(* IEC 61131-3 sources: daoli-st-library/DL_Process (part 68) *)

(* ---- FB_DL_MultiZoneSetpointScheduler.st ---- *)
(*==============================================================================
 * 组件名称 (Component)  : FB_DL_MultiZoneSetpointScheduler
 * 所属子库 (Sublibrary) : DL_Process ｜ 版本 (Version) : 1.0.2 ｜ 2026-11-23
 * 兼容性   (Platform)   : CODESYS 3.5+ / TwinCAT 3 / 汇川 InoProShop / 施耐德 Machine Expert
 *                         仅依赖 IEC 61131-3 标准（FOR / CASE / ABS），零厂商私有库
 * 功能描述 (Function)   : 多区设定值按时段表切换（4 区 × 每区最多 8 时段）。每区持有一张
 *                         「起始分钟 + 设定值」时段表，按当日第几分钟 nMinuteOfDay 选出生效
 *                         时段，并把「与上一生效值不同」的区以 abSpChanged 单拍沿上报。
 *                         参数非法（时段非单调 / 分钟越域 / 设定值非有限 / 时段数越界）→
 *                         整机进 eFault 并锁存首个成因码；eFault 唯一出口为 bReset（重校验通过）。
 *                         **时钟来源声明**：本件不读任何系统时钟（零全局耦合 R1），
 *                         nMinuteOfDay 由上层 PRG 从 RTC 换算后传入（0..1439）。
 *                         **bEnable = FALSE 语义（R191 二选一，本件选「冻结保持末值」）**：
 *                         各区 afActiveSp / aiActiveIdx 保持末值不动，abSpChanged 不再发沿，
 *                         bValid 落 FALSE 提示「该值已不与时钟对齐」。
 * 接口     (Interface)  : 输入 bEnable / bReset / nMinuteOfDay / aiZoneSlotCount[1..4] /
 *                         aSlots[1..4][1..8]（ST_DL_SpSlot）；输出 afActiveSp[1..4] /
 *                         aiActiveIdx[1..4] / abSpChanged[1..4]（单拍）/ eState / bError /
 *                         eCause / bValid / nFaultZone。
 * 状态迁移表 (State Transition Table)：
 *   ① eIdle → eApply：bEnable 上升（或上电首拍 bEnable 已为 TRUE）；
 *      拍 N 进入（bEnable 为 TRUE）/ 本拍行为：不做选段、不发沿、冻结保持 / 拍 N+1 转出至 eApply。
 *      拒收：bEnable 为 FALSE 时本拍不迁出，abSpChanged 保持 FALSE。
 *   ② eApply → eHold：全量参数校验通过且选段、比对、发沿完成（同一拍内完成）；
 *      拍 N 进入（校验通过）/ 本拍行为：写出 afActiveSp/aiActiveIdx 与 abSpChanged 单拍沿 /
 *      拍 N+1 转出至 eHold。
 *   ③ eApply → eFault：任一区校验失败（时段数越界 / 分钟越域 / 时段非单调 / 设定值非有限）；
 *      拍 N 进入（校验失败）/ 本拍行为：锁存首个成因码、不写 afActiveSp（保持末值）/
 *      拍 N+1 转出至 eFault（段尾迁移闸）。
 *   ④ eHold → eApply：nMinuteOfDay 落在任一时段起点（时段边界）或 bReset 为 TRUE（强制重校验）；
 *      拍 N 进入（边界命中或复位）/ 本拍行为：交出控制权、本拍不写设定值 / 拍 N+1 转出至 eApply。
 *   ⑤ eHold → eIdle：bEnable 落 FALSE（失能退出，出口冻结保持）。
 *   ⑥ eHold → eFault：段尾迁移闸（锁存位已置）——由①②③④ 任一分支置锁存后同拍迁入。
 *   ⑦ eFault → eIdle：bReset 上升且 NOT bEnable（复位沿要求先失能，避免带故障参数直接投产）；
 *      拍 N 进入（bReset 沿 + 已失能）/ 本拍行为：清锁存与成因码 / 拍 N+1 转出至 eIdle。
 *      该路径可达性自证：bReset 与 bEnable 均为外部引脚，恒可到达（R152）。
 *   ⑧ ELSE（非法枚举值）→ eFault，成因码 eIllegalState（R6 兜底）。
 * 边界     (Boundary)   : ① 首时段之前（nMinuteOfDay < 第 1 段起始）：取第 1 段值（日头承接），
 *                            该口径在段 4 注释内声明，不置码。
 *                         ② nMinuteOfDay 越域（<0 或 >1439）→ 钳位到 [0,1439] 并置信息级
 *                            eMinuteClamped（信息级永不置 bError）。
 *                         ③ 数组下标访问前先以 nCnt ∈ [1,8] 钳定（R4），越界槽不访问。
 *                         ④ 浮点同值比较用容差 DL_MZS_EPS（1E-6），禁 `=`（R4）。
 *                         ⑤ 零全局耦合（无 GVL / VAR_EXTERNAL / %I / %Q）。
 * 码表     (Codes)      : 本件不占用全局数字码位（R297 零码位范式）；出口为 BOOL + ENUM，
 *                         enum E_DL_MzsCause 归属本文件（全库唯一属主）。信息级
 *                         eMinuteClamped / eNoChange 永不置 bError；故障级成因码各占独立成员
 *                         （R190 归因唯一），锁存回放至 bReset 沿（FB33-1）。
 * 分工声明 (Scope)      : 时段选择与下发归本件；设定值斜坡 / 无扰切换归 FB_DL_RampGenerator 类；
 *                         PID 闭环归温控件。本件不下装任何硬件输出。
 * 归属     (Ownership)  : E_DL_MzsState / E_DL_MzsCause / ST_DL_SpSlot 归属本文件
 *                         （全库唯一定义，R264），引用件只引用不重声明。
 * 红线自检 (Redline)    : R1 ✓ 零 GVL ｜ R2 ✓ 零 %I/%Q ｜ R3 ✓ 纯 IEC ｜ R4 ✓ 下标钳定 +
 *                         非有限双判 + 容差比较 + 循环界固定 ｜ R5 ✓ 逐行同行双语注释
 *                         R6 ✓ 四态 ENUM + CASE + ELSE ｜ R7 N/A（本件无需定时器/边沿实例）
 *                         R14 ✓ 无 PROPERTY ｜ R8/R9 N/A（无 METHOD）
 * 修订历史 (Revision)   : 2026-11-24  v1.0.2  R79-F2/P3：bReset 电平→R_TRIG 沿 + eHold 复位沿同步清锁存（原头版本号滞留 1.0.0，已核正）
 *                         2026-11-23  v1.0.0  R78-B3 首版
 *                         2026-11-23  v1.0.1  R78 返修：E045 数组访问改嵌套索引形式（8 处）；
 *                                             eHold 相补时段数重校验闸（越界锁存 eBadCount）；
 *                                             M5：成功路径不再覆盖钳位信息级码
 * 验收向量 (Acceptance) :
 *   V1 bEnable=TRUE、nMinuteOfDay=480、区 1 时段表 {(0,20.0),(480,22.0)} → afActiveSp[1]=22.0,
 *      aiActiveIdx[1]=2, abSpChanged[1]=TRUE 单拍；次拍 abSpChanged[1]=FALSE。
 *   V2 续 V1、nMinuteOfDay 保持 481（非边界）→ eState=eHold，无沿。
 *   V3 区 2 时段表起始分钟 {0, 600, 500}（非单调）→ eState=eFault, eCause=eSlotNotMonotonic,
 *      bError=TRUE, afActiveSp[2] 保持末值；bReset 上升且 bEnable=FALSE → 回 eIdle。
 *   V4 nMinuteOfDay=2000（越域）→ 钳位到 1439，eCause=eMinuteClamped（信息级），bError=FALSE。
 *   V5 区 3 设定值为 NaN → eState=eFault, eCause=eBadSetpoint, bError=TRUE。
 *============================================================================*)

(*-----------------------------------------------------------------------------
 * 结构体: ST_DL_SpSlot（时段表行：起始分钟 + 该时段设定值），归属本文件，全库唯一属主
 *----------------------------------------------------------------------------*)
TYPE ST_DL_SpSlot :
STRUCT
    nStartMin : INT := 0;      // 时段起始时刻（当日第几分钟，0..1439）[-] / Slot start minute of the day
    fSetpoint : REAL := 0.0;   // 该时段生效设定值 [工程单位，由调用方标定] / Setpoint effective within the slot
END_STRUCT
END_TYPE

(*-----------------------------------------------------------------------------
 * 枚举: E_DL_MzsState（状态机相位；eFault 为安全相，仅 bReset 沿迁出）
 *----------------------------------------------------------------------------*)
TYPE E_DL_MzsState :
(
    eIdle  := 0,    // 空闲：未使能，设定值冻结保持末值 / Idle: disabled, setpoints frozen at last value
    eApply := 10,   // 校验与应用：全量参数校验 + 选段 + 比对 + 发沿（同拍完成）/ Validate and apply in one scan
    eHold  := 20,   // 驻留：等时段边界或复位，每拍只做边界检测 / Hold: wait for a slot boundary or reset
    eFault := 90    // 故障安全相：参数非法，锁存成因码，仅 bReset 沿迁出 / Fault latched, reset edge only
);
END_TYPE

(*-----------------------------------------------------------------------------
 * 枚举: E_DL_MzsCause（成因码；信息级 = 0..9，故障级 = 10 起，各成因独立成员 R190）
 *----------------------------------------------------------------------------*)
TYPE E_DL_MzsCause :
(
    eNone             := 0,   // 信息级：无事件 / Info: no event
    eMinuteClamped    := 1,   // 信息级：当日分钟越域已钳位 / Info: minute of day clamped into range
    eSlotNotMonotonic := 10,  // 故障级：时段起始分钟非严格递增 / Fault: slot start minutes not strictly increasing
    eBadMinute        := 11,  // 故障级：单条时段起始分钟越域 / Fault: slot start minute out of range
    eBadCount         := 12,  // 故障级：时段数越界（不在 1..8）/ Fault: slot count out of the 1..8 range
    eBadSetpoint      := 13,  // 故障级：设定值非有限 / Fault: non-finite setpoint
    eIllegalState     := 14   // 故障级：非法状态枚举值（CASE ELSE 兜底）/ Fault: illegal state enum value
);
END_TYPE

FUNCTION_BLOCK FB_DL_MultiZoneSetpointScheduler
VAR_INPUT
    bEnable        : BOOL := FALSE;                       // 使能：FALSE 冻结保持末值（本件语义声明）/ Enable, FALSE freezes the last setpoints
    bReset         : BOOL := FALSE;                       // 复位（上升沿）：清故障锁存并要求失能 / Reset rising edge clears the fault latch and requires disabled state
    nMinuteOfDay   : INT := 0;                            // 当日第几分钟，有效域 0..1439 [-] / Minute of the day, valid domain 0..1439
    aiZoneSlotCount : ARRAY[1..4] OF INT;                 // 各区时段条数，有效域 1..8 [-] / Slot count per zone, valid domain 1..8
    aSlots         : ARRAY[1..4] OF ARRAY[1..8] OF ST_DL_SpSlot;  // 四区 × 八时段时段表 / Slot tables of four zones with up to eight slots each
END_VAR
VAR_OUTPUT
    afActiveSp  : ARRAY[1..4] OF REAL;      // 各区当前生效设定值（冻结保持，见 bEnable 语义）[工程单位] / Active setpoint per zone
    aiActiveIdx : ARRAY[1..4] OF INT;       // 各区当前生效时段序号（1..8），未选定时为 0 [-] / Active slot index per zone
    abSpChanged : ARRAY[1..4] OF BOOL;      // 各区设定值变更单拍沿（统一出口预置，FB51-8）[-] / Single-scan change flag per zone
    eState      : E_DL_MzsState;            // 状态出口（段尾单点映射）[-] / State outlet, mapped at the tail
    bError      : BOOL;                     // 故障锁存标志（仅故障级成因置位）[-] / Fault latch flag
    eCause      : E_DL_MzsCause;            // 成因码出口（锁存回放）[-] / Cause code outlet, replayed from the latch
    bValid      : BOOL;                     // 设定值有效回执（eHold 且参数有效才 TRUE）[-] / Setpoint validity receipt
    nFaultZone  : INT;                      // 首个故障所在区号（0 = 无故障 / 全局性故障）[-] / Zone index of the first fault
END_VAR
VAR
    _eState      : E_DL_MzsState := E_DL_MzsState.eIdle;   // 内部相位（CASE 唯一写入目标）[-] / Internal phase
    _bFaultLatch : BOOL := FALSE;                          // 故障锁存位（仅 bReset 沿清除）[-] / Fault latch bit cleared by the reset edge only
    _eCauseLatch : E_DL_MzsCause := E_DL_MzsCause.eNone;    // 锁存成因码（锁存回放，FB33-1）[-] / Latched cause code replayed to the outlet
    _nFaultZone  : INT := 0;                               // 首个故障区号 [1..4]，0 表示无 / Zone index of the first fault
    _bParamOk    : BOOL := TRUE;                           // 本拍参数校验通过标志 [-] / Parameter validation flag of this scan
    _eCauseTmp   : E_DL_MzsCause := E_DL_MzsCause.eNone;    // 本拍首个成因（未锁存）[-] / First cause of this scan before latching
    _nFaultZtmp  : INT := 0;                               // 本拍首个故障区号（未锁存）[-] / First fault zone of this scan before latching
    _nMinute     : INT := 0;                               // 钳位后的当日分钟 [0..1439] / Clamped minute of the day
    _nCnt        : INT := 0;                               // 当前区时段条数（校验后使用）[-] / Slot count of the current zone
    _nIdx        : INT := 0;                               // 选段中间结果（时段序号）[-] / Intermediate slot index
    _nNewIdx     : INT := 0;                               // 本区本拍应生效时段序号 [-] / Slot index that should be active this scan
    _fNewSp      : REAL := 0.0;                            // 本区本拍应生效设定值 [工程单位] / Setpoint that should be active this scan
    _bBoundary   : BOOL := FALSE;                          // 时段边界命中标志（eHold 用）[-] / Slot boundary hit flag used in eHold
    _nZ          : INT := 0;                               // 外层循环索引：区号 [1..4] / Outer loop index, zone number
    _nK          : INT := 0;                               // 内层循环索引：时段序号 [1..8] / Inner loop index, slot number
    _rtReset     : R_TRIG;                                 // 复位沿检测实例（v1.0.1 补：声明沿即实现沿，段 1 无条件刷新）/ Reset edge detector, refreshed unconditionally in segment 1
END_VAR
VAR CONSTANT
    DL_MZS_ZONES    : INT := 4;             // 固定区数（数组第一维上界）[-] / Fixed zone count, upper bound of dimension one
    DL_MZS_SLOTS    : INT := 8;             // 每区最大时段数（数组第二维上界）[-] / Max slots per zone, upper bound of dimension two
    DL_MZS_MIN_DAY  : INT := 1439;          // 当日最大分钟数（23:59）[-] / Last minute of the day
    DL_MZS_MIN_ONE  : INT := 1;             // 时段数下界 [-] / Lower bound of the slot count
    DL_MZS_ZERO     : INT := 0;             // 整数零基准 [-] / Integer zero base
    DL_MZS_FZERO    : REAL := 0.0;          // 实数零基准 [-] / Real zero base
    DL_MZS_EPS      : REAL := 1.0E-6;       // 设定值同值判定容差 [-] / Setpoint equality tolerance
    DL_MZS_FIN      : LREAL := 1.0E308;     // 有限性判据上界（R477：ABS(x)>FIN 判 Inf）[工程单位] / finiteness ceiling flags Inf
END_VAR

(* —— 段 1：单拍位与当拍工作量预置（只清单拍标志，不清锁存/保持量，FB32-1） —— *)
_rtReset(CLK := bReset);                                // 复位沿刷新必须无条件周期调用（R7；v1.0.1 修复 J1 电平判据缺陷）/ The reset edge must be refreshed unconditionally every scan
FOR _nZ := 1 TO DL_MZS_ZONES DO
    abSpChanged[_nZ] := FALSE;                          // 变更沿每拍先预清 / Change edge preset FALSE every scan
END_FOR
_bParamOk   := TRUE;                                    // 校验标志复位 / Validation flag reset
_eCauseTmp  := E_DL_MzsCause.eNone;                      // 当拍成因复位 / Scan cause reset
_nFaultZtmp := DL_MZS_ZERO;                             // 当拍故障区复位 / Scan fault zone reset
_bBoundary  := FALSE;                                   // 边界标志复位 / Boundary flag reset
eCause      := E_DL_MzsCause.eNone;                      // 成因出口每拍预置信息级零码（段 2/段 3 内改写）/ Cause outlet preset to the info zero code every scan

(* —— 段 2：入参钳位与域闸（分钟越域钳位并置信息级，R4 下标与域安全） —— *)
_nMinute := nMinuteOfDay;                               // 取入参 / Take the input pin
IF _nMinute < DL_MZS_ZERO THEN
    _nMinute  := DL_MZS_ZERO;                           // 下越界钳到 0 / Clamp low
    eCause    := E_DL_MzsCause.eMinuteClamped;          // 信息级：已钳位 / Info: clamped
ELSIF _nMinute > DL_MZS_MIN_DAY THEN
    _nMinute  := DL_MZS_MIN_DAY;                        // 上越界钳到 1439 / Clamp high
    eCause    := E_DL_MzsCause.eMinuteClamped;          // 信息级：已钳位 / Info: clamped
END_IF

(* —— 段 3：状态机主体（唯一相位写入点，每分支迁移条件自足） —— *)
CASE _eState OF
    E_DL_MzsState.eIdle :
        (* 迁移①：使能上升进入统一校验相；未使能则保持冻结语义 *)
        IF bEnable THEN
            _eState := E_DL_MzsState.eApply;            // 迁入校验与应用相 / Move to validate-and-apply
        END_IF

    E_DL_MzsState.eApply :
        IF NOT bEnable THEN
            _eState := E_DL_MzsState.eIdle;             // 使能消失：退回冻结 / Enable gone: back to idle
        ELSE
            (* 段 4 前置：逐区全量校验（时段数 → 单条分钟 → 单调性 → 设定值有限性） *)
            FOR _nZ := 1 TO DL_MZS_ZONES DO
                _nCnt := aiZoneSlotCount[_nZ];          // 取本区时段条数 / Slot count of this zone
                IF (_nCnt < DL_MZS_MIN_ONE) OR (_nCnt > DL_MZS_SLOTS) THEN
                    _bParamOk := FALSE;                 // 时段数越界 / Count out of range
                    IF _eCauseTmp = E_DL_MzsCause.eNone THEN
                        _eCauseTmp  := E_DL_MzsCause.eBadCount;    // 首因锁存用 / First cause kept
                        _nFaultZtmp := _nZ;                        // 记录故障区号 / Record the fault zone
                    END_IF
                ELSE
                    FOR _nK := 1 TO _nCnt DO
                        (* 单条起始分钟域闸：0..1439 *)
                        IF (aSlots[_nZ][_nK].nStartMin < DL_MZS_ZERO)
                            OR (aSlots[_nZ][_nK].nStartMin > DL_MZS_MIN_DAY) THEN
                            _bParamOk := FALSE;
                            IF _eCauseTmp = E_DL_MzsCause.eNone THEN
                                _eCauseTmp  := E_DL_MzsCause.eBadMinute;   // 故障级：分钟越域
                                _nFaultZtmp := _nZ;
                            END_IF
                        END_IF
                        (* 单调性闸：自第 2 条起必须严格大于前一条 *)
                        IF _nK > 1 THEN
                            IF aSlots[_nZ][_nK].nStartMin <= aSlots[_nZ][_nK - 1].nStartMin THEN
                                _bParamOk := FALSE;
                                IF _eCauseTmp = E_DL_MzsCause.eNone THEN
                                    _eCauseTmp  := E_DL_MzsCause.eSlotNotMonotonic;   // 故障级：非单调
                                    _nFaultZtmp := _nZ;
                                END_IF
                            END_IF
                        END_IF
                        (* 设定值有限性闸（R79 双判） *)
                        (* v1.0.2 补（闸 Q2）：Inf 判据改 R477 范式 ABS(x) > DL_MZS_FIN，
                           x−x 差判在部分编译器会常量折叠成 0，Inf 设定值可穿透写入 afActiveSp *)
                        IF (aSlots[_nZ][_nK].fSetpoint <> aSlots[_nZ][_nK].fSetpoint)
                            OR (ABS(aSlots[_nZ][_nK].fSetpoint) > DL_MZS_FIN) THEN
                            _bParamOk := FALSE;
                            IF _eCauseTmp = E_DL_MzsCause.eNone THEN
                                _eCauseTmp  := E_DL_MzsCause.eBadSetpoint;   // 故障级：设定值非有限
                                _nFaultZtmp := _nZ;
                            END_IF
                        END_IF
                    END_FOR
                END_IF
            END_FOR

            IF NOT _bParamOk THEN
                (* 迁移③：校验失败 → 锁存首因（不改写 afActiveSp，保持末值） *)
                _eCauseLatch := _eCauseTmp;                 // 锁存成因码 / Latch the cause code
                _nFaultZone  := _nFaultZtmp;                // 锁存故障区号 / Latch the fault zone
                _bFaultLatch := TRUE;                       // 置故障锁存（段尾迁移闸迁相）/ Latch the fault
            ELSE
                (* 段 4：选段 + 比对 + 发沿（每区独立裁决，日头承接口径见分支注释） *)
                FOR _nZ := 1 TO DL_MZS_ZONES DO
                    _nCnt   := aiZoneSlotCount[_nZ];        // 时段条数 / Slot count
                    _nNewIdx := DL_MZS_MIN_ONE;             // 缺省取第 1 段（日头承接：首段之前沿用首段值）/ Default first slot
                    FOR _nK := 1 TO _nCnt DO
                        IF aSlots[_nZ][_nK].nStartMin <= _nMinute THEN
                            _nNewIdx := _nK;                // 最后一条不晚于当前分钟的时段生效 / Last slot not later than now wins
                        END_IF
                    END_FOR
                    _fNewSp := aSlots[_nZ][_nNewIdx].fSetpoint;    // 取该时段设定值 / Setpoint of the winning slot
                    IF (ABS(afActiveSp[_nZ] - _fNewSp) >= DL_MZS_EPS) OR (aiActiveIdx[_nZ] <> _nNewIdx) THEN
                        afActiveSp[_nZ]  := _fNewSp;            // 写入生效设定值 / Write the active setpoint
                        aiActiveIdx[_nZ] := _nNewIdx;           // 写入生效时段序号 / Write the active slot index
                        abSpChanged[_nZ] := TRUE;               // 单拍变更沿（本拍置位，次拍段 1 预清）/ Single-scan change edge
                    END_IF
                END_FOR
                IF eCause <> E_DL_MzsCause.eMinuteClamped THEN
                    eCause := E_DL_MzsCause.eNone;          // 信息级：无事件（M5：不覆盖段 2 已置的钳位信息码）/ Info: no event, keep the pre-set clamp code
                END_IF
                _bFaultLatch := FALSE;                      // 校验通过：清故障锁存（正常路径唯一清点）/ Clear the latch on the valid path
                _eState := E_DL_MzsState.eHold;             // 迁移②：进入驻留相 / Move to hold
            END_IF
        END_IF

    E_DL_MzsState.eHold :
        IF NOT bEnable THEN
            _eState := E_DL_MzsState.eIdle;                 // 迁移⑤：失能退出（冻结保持）/ Disable exit, frozen
        ELSE
            (* 边界检测：任一时段起点等于当前分钟（或日切 0 点）→ 回校验相重算 *)
            IF _nMinute = DL_MZS_ZERO THEN
                _bBoundary := TRUE;                         // 日切 0 点视为边界 / Day roll-over counts as a boundary
            END_IF
            FOR _nZ := 1 TO DL_MZS_ZONES DO
                _nCnt := aiZoneSlotCount[_nZ];              // 取本区时段条数（引脚每拍可被外部改写，不信任 eApply 旧校验）/ Slot count, pin may change every scan
                IF (_nCnt < DL_MZS_MIN_ONE) OR (_nCnt > DL_MZS_SLOTS) THEN
                    (* L1 加固：eHold 相重校验失败 → 故障锁存（复用参数校验闸同款 eBadCount），跳出该区处理 *)
                    IF _eCauseLatch = E_DL_MzsCause.eNone THEN   // 首因保留（不覆盖既有锁存码）/ Keep the first cause
                        _eCauseLatch := E_DL_MzsCause.eBadCount; // 故障级：时段数越界（既有成因成员，R190）/ Fault: count out of range
                        _nFaultZone  := _nZ;                     // 锁存故障区号 / Latch the fault zone
                    END_IF
                    _bFaultLatch := TRUE;                        // 置故障锁存（段 5 迁移闸同拍迁入 eFault）/ Latch the fault
                ELSE
                    FOR _nK := 1 TO _nCnt DO
                        IF aSlots[_nZ][_nK].nStartMin = _nMinute THEN
                            _bBoundary := TRUE;                 // 时段边界命中 / Slot boundary hit
                        END_IF
                    END_FOR
                END_IF
            END_FOR
            IF _rtReset.Q THEN
                (* v1.0.2 补（闸 P3）：eHold 内复位沿属"强制重校验"语义，必须同时清故障锁存，
                   否则 eApply 重校验通过后 bError 仍为 TRUE（声明"复位即清锁存"未兑现） *)
                _bFaultLatch := FALSE;                      // 复位沿清故障锁存 / Reset edge clears the fault latch
                _eCauseLatch := E_DL_MzsCause.eNone;        // 复位沿清锁存成因 / Reset edge clears the latched cause
                eCause       := E_DL_MzsCause.eNone;        // 出口同步归零 / Outlet follows
                nFaultZone   := DL_MZS_ZERO;                // 故障区号归零 / Fault zone index cleared
            END_IF
            IF (NOT _bFaultLatch) AND (_bBoundary OR _rtReset.Q) THEN
                _eState := E_DL_MzsState.eApply;            // 迁移④：边界命中或强制重校验（R274：锁存期禁迁入执行相）/ Boundary or forced revalidation
            END_IF
        END_IF

    E_DL_MzsState.eFault :
        (* 迁移⑦：唯一出口 —— bReset 沿 + 已失能（避免带故障参数直接投产） *)
        IF _rtReset.Q AND (NOT bEnable) THEN
            _bFaultLatch := FALSE;                          // 清故障锁存 / Clear the fault latch
            _eCauseLatch := E_DL_MzsCause.eNone;            // 清锁存成因 / Clear the latched cause
            _nFaultZone  := DL_MZS_ZERO;                    // 清故障区号 / Clear the fault zone
            _eState      := E_DL_MzsState.eIdle;            // 回空闲相 / Back to idle
        END_IF

ELSE
    (* 迁移⑧：非法枚举值兜底（R6） *)
    _eCauseLatch := E_DL_MzsCause.eIllegalState;            // 故障级：非法状态 / Fault: illegal state value
    _bFaultLatch := TRUE;                                   // 置锁存 / Latch
    _eState      := E_DL_MzsState.eFault;                   // 迁入安全相 / Move to the safe state
END_CASE

(* —— 段 5：段尾故障迁移闸（FB50-1④：锁存与迁相分离，置于解除段之后） —— *)
IF _bFaultLatch AND (_eState <> E_DL_MzsState.eFault) THEN
    _eState := E_DL_MzsState.eFault;                        // 锁存即迁相 / Latch forces the fault phase
END_IF

(* —— 段 6：统一出口（状态映射 + 锁存回放 + 单拍位已由段 1 预置） —— *)
eState := _eState;                                          // 相位映射 / Phase mapping
bError := _bFaultLatch;                                     // 故障标志取锁存位（派生式）/ Fault flag derived from the latch
IF _bFaultLatch THEN
    eCause := _eCauseLatch;                                 // 故障期回放锁存码（FB33-1）/ Replay the latched code
    nFaultZone := _nFaultZone;                              // 回放故障区号 / Replay the fault zone
ELSE
    nFaultZone := DL_MZS_ZERO;                              // 无故障：区号归零 / No fault: zone index zero
END_IF
bValid := (_eState = E_DL_MzsState.eHold) AND (NOT _bFaultLatch);   // 仅驻留相且无锁存时值可信 / Valid only in hold without a latch
END_FUNCTION_BLOCK

(* ---- FB_DL_OccScheduleWindow.st ---- *)
(*==============================================================================
 * 组件名称 (Component)  : FB_DL_OccScheduleWindow
 * 所属子库 (Sublibrary) : DL_Process
 * 当前版本 (Version)    : 1.0.0
 * 组件分类 (Category)   : 功能块（FUNCTION_BLOCK）· 多窗作息排程 ·
 *                         Level 2 行业池 9.5 节 P0 链路闭环示范
 * 兼容性   (Platform)   : CODESYS 3.5 / TwinCAT 3 / 汇川 InoProShop / Schneider
 *                         Machine Expert；仅依赖 Standard.library（R_TRIG /
 *                         MIN）与本库 DL_Base 已入库组件，零厂商方言
 * 功能描述 (Function)   : 多窗作息排程块（最多 4 窗并行）。日期/时刻全部引脚
 *                         注入（零全局耦合红线：禁读 CPU 本地钟）→ 调用
 *                         FC_DL_DayOfWeekCalc 换算当日星期（ISO-8601 序）
 *                         → 内部 4 实例复用 FB_DL_TimeWindowCheck 逐窗判定
 *                         （每日窗矩阵 + 节假日覆盖位）→ 输出占用合成、
 *                         占用开始沿单发、活动窗号（多窗同开取最小号）与
 *                         预启动占位（提前启机预热/预冷用）。
 * 设计要点 (Key notes)  : ① 每窗占用 = 窗实例 bInWindow（内部已合成 总使能
 *                           AND 星期位 AND 时刻窗），总使能引脚折入
 *                           bEnableDay := aWinEnable[i] AND NOT aHoliday-
 *                           Override[i]（节假日强制当日该窗关闭）；窗实例的
 *                           aWeekdayEnable 由本块按 aWeekdayWin[i, 当日星期]
 *                           单日位展开为 7 日表填充；
 *                         ② 预启动占位：折算「占用开始时刻 − tPreLeadTime」
 *                           分钟域判定。推导：窗开始分钟 uStartMin（UINT 域，
 *                           0..1439，与 FB_DL_TimeWindowCheck 折算口径一致）；
 *                           当 提前量 ≤ 开始时刻 时预启带 = [开始−提前, 开始)
 *                           （左闭右开）；当 提前量 > 开始时刻（跨零点回绕）
 *                           时预启带 = [开始+24h−提前, 开始)∪[0, 开始)，即
 *                           [开始+1440−lead, 1440) 与 [0, 开始) 的并——本块
 *                           统一用 TIME 域表达（T#24H 回绕式），时刻折算先
 *                           USINT→DINT 扩宽再乘 60 防溢出（复用窗实例口径，
 *                           声明一致）；预启带归属注入日期当日窗（跨零点前段
 *                           归属前一日期的同一窗组态，调用方按日切换注入即可）；
 *                         ③ 窗实例与沿检测实例在主体无条件周期刷新（R7，
 *                           严禁置于 IF/CASE 分支）；
 *                         ④ 【事件型+日切换沿，免首扫（R23）】输入输出均为
 *                           电平/日历注入，无连续量同步语义，窗判定为组合
 *                           逻辑逐拍重算，故不设 bInit 首扫判据；
 *                         ⑤ 日期越界（FC 返回 eInvalid）→ 全窗按不在窗处理
 *                           + 信息级 0005_0210；各窗实例信息级码 0001_0202
 *                           不透传，本块归并为自身码 0005_0211（头注释声明）；
 *                         ⑥ bReset 上升沿清除当拍信息级码（日切换后防陈旧码
 *                           残留），不影响窗判定结果（沿用窗实例 D2 语义）；
 *                         ⑦ 本块无浮点量，非有限值防御不适用（公约 0.8 N/A）。
 * 枚举归属 (Enum note)  : 复用 E_DL_Weekday（DL_Base，随 FC_DL_DayOfWeekCalc
 *                         同文件发布的既有公开契约，直接引用，禁止重定义）；
 *                         本块不新增任何 DUT。
 * 依赖     (Depends)    : FB_DL_TimeWindowCheck（DL_Base，4 实例复用）；
 *                         FC_DL_DayOfWeekCalc + E_DL_Weekday（DL_Base）；
 *                         Standard.library：R_TRIG / MIN。
 * 开源溯源 (Origin)     : 原创实现（参考 OSCAT Building 时钟排程族与
 *                         Siemens LGF 定时开关族的公开行为定义，clean-room）。
 *                         仅借鉴「多窗排程 + 星期使能矩阵 + 节假日覆盖」的
 *                         公开行为语义；多实例单一语义组合架构、预启动占位、
 *                         时间引脚注入均为本库独立设计，未复制任何源码行。
 * 故障码表 (Error codes):
 *   16#0005_0210【信息级】日期参数越界（年/月/日，FC 返回 eInvalid），全窗
 *                 按不在窗处理
 *   16#0005_0211【信息级】窗时刻参数越界（各窗实例 0001_0202 码不透传，本块
 *                 归并为自身码；实例侧越界已钳位照常计算，本块预启动判定对
 *                 参数越界窗按跳过处理）
 *   【02xx 段信息级占位声明（规格 §7 有意裁定，R11 留档）】0210/0211 占用
 *   02xx 段：日历排程块全部事件均为信息级（无安全联锁、无锁存故障位），
 *   故障级段整体保留给后续工艺联锁件，沿用 FB_DL_TimeWindowCheck 先例，
 *   避免读者误判为故障级。
 * 红线自检 (Redline)    : R1 ✓ 零全局变量表与外部变量引用 ｜ R2 ✓ 零物理 IO 地址直写
 *                         R3 ✓ 纯 IEC 61131-3 ｜ R4 ✓ 数组索引域校验+USINT→DINT
 *                             扩宽防溢出+TIME 回绕防御（提前量钳位）；无浮点量，
 *                             非有限值防御不适用（R23 事件型）
 *                         R5 ✓ 全变量中英双语同行注释
 *                         R6 不适用（组合逻辑+沿检测，无状态机；星期换算
 *                           CASE 含 ELSE 兜底）
 *                         R7 ✓ 4 个窗实例 + 2 个 R_TRIG 实例主体无条件周期刷新
 * 修订历史 (Revision)   :
 *   2026-11-15  v1.0.0  首版入库 · Round 06 · 泳道 C · 契约出处 ROUND_PLAN_R6 §3.15
 * 验收向量 (Acceptance) :
 *   V1 单窗占用链：窗 1 On=08:00/Off=18:00 使能，Now=07:59 → bOccupied=
 *      FALSE；08:00 当拍 bPulseOnOccupy=TRUE 单发且 bOccupied=TRUE；
 *      18:00 当拍 bOccupied=FALSE（左闭右开与窗实例一致）
 *   V2 四窗并行：窗 2 与窗 4 同时在窗 → uActiveWin=2（多窗同开取最小号）
 *   V3 节假日覆盖：aHolidayOverride[1]=TRUE → 当日窗 1 强制不在窗，其余窗
 *      不受影响
 *   V4 预启动提前量（含跨零点回绕）：tPreLeadTime=T#30M，窗 On=06:00 →
 *      Now=05:35 bPreStart=TRUE 且 bOccupied=FALSE，06:00 当拍 bPreStart
 *      随占用置位而清零；跨零点窗 On=00:10、提前量 30 分 → Now=23:50 时
 *      bPreStart=TRUE（预启带 [23:40, 00:10)，回绕式 开始+24h−提前=23:40）
 *   V5 日期越界降级：uMonth=13 → FC 返回 eInvalid → 全窗不在窗 +
 *      0005_0210；bReset 沿当拍清码
 *   V6 星期矩阵按日生效：aWeekdayWin[1,6]=FALSE（周六位）→ 周六窗 1 不在窗，
 *      周一~周五正常
 *============================================================================*)

(*-----------------------------------------------------------------------------
 * 调用示例 (Instance guide)：
 *   fbOcc.uYear := 2026; fbOcc.uMonth := 11; fbOcc.uDay := 15;   // 日历注入
 *   fbOcc.uHourNow := stClock.hour; fbOcc.uMinNow := stClock.min;
 *   fbOcc.aWinEnable[1] := TRUE; fbOcc.aHourOn[1] := 8;         // 窗 1 组态，其余 3 窗同构
 *   fbOcc(tPreLeadTime := T#30M, bReset := bDaySwReset);         // 周期调用
 *   预热/预冷联动：bPreStart → AHU 通风预启（非占用占位）；bPulseOnOccupy
 *   → 占用开始沿一次性事件（照明/门禁联动）。uActiveWin 供 HMI 显示当前窗。
 *----------------------------------------------------------------------------*)

FUNCTION_BLOCK FB_DL_OccScheduleWindow
VAR_INPUT
    uYear              : UINT;             // 日期注入-年（Injected date year）[年] 有效域 1980..2099，越界返回 eInvalid（透传 FC_DL_DayOfWeekCalc）
    uMonth             : USINT;            // 日期注入-月（Injected month）[月] 有效域 1..12，越界按日期非法处理
    uDay               : USINT;            // 日期注入-日（Injected day）[日] 有效域 1..当月天数（含闰年），越界按日期非法处理
    uHourNow           : USINT;            // 当前时刻注入-时（Injected time hour）[h] 0..23，越界按不在窗处理（禁读 CPU 钟，公约 0.9）
    uMinNow            : USINT;            // 当前时刻注入-分（Injected time minute）[min] 0..59
    aWinEnable         : ARRAY[1..4] OF BOOL;          // 各窗使能（Window enables）[1] 窗 1..4，FALSE 时该窗恒不在窗
    aHourOn            : ARRAY[1..4] OF USINT;         // 各窗开启时刻-时（Window on hours）[h] 0..23，越界该窗预启动跳过（实例侧钳位照算）
    aMinOn             : ARRAY[1..4] OF USINT;         // 各窗开启时刻-分（Window on minutes）[min] 0..59
    aHourOff           : ARRAY[1..4] OF USINT;         // 各窗关闭时刻-时（Window off hours）[h] 0..23，支持跨零点窗
    aMinOff            : ARRAY[1..4] OF USINT;         // 各窗关闭时刻-分（Window off minutes）[min] 0..59
    aWeekdayWin        : ARRAY[1..4, 1..7] OF BOOL;    // 各窗星期使能矩阵（Per-window weekday matrix）[1] 第二维 1=周一..7=周日（ISO 序）
    aHolidayOverride   : ARRAY[1..4] OF BOOL;          // 节假日覆盖位（Holiday overrides）[1] TRUE=当日该窗强制关闭
    tPreLeadTime       : TIME := T#30M;    // 预启动提前量（Pre-start lead time）默认 T#30M，防御钳位 ≤ T#12H，占用开始前输出预启动占位
    bReset             : BOOL := FALSE;    // 复位（Reset）[1] 上升沿：清除当拍信息级码（不影响窗判定）
END_VAR
VAR_OUTPUT
    bOccupied          : BOOL;             // 占用中（Occupied）[1] 任一有效窗在窗内
    bPreStart          : BOOL;             // 预启动占位（Pre-start placeholder）[1] 未占用且距某有效窗开始 ≤ 提前量
    bPulseOnOccupy     : BOOL;             // 占用开始沿单发（Occupancy start edge）[1] TRUE 持续一拍
    uActiveWin         : USINT;            // 当前活动窗号（Active window index）1..4，0=无，多窗同开取最小号
    uErrorId           : UDINT;            // 信息级码（Info code）16#0005_0210 日期非法 / 16#0005_0211 窗参数越界；0 = 无
END_VAR
VAR
    _fbWin1            : FB_DL_TimeWindowCheck;  // 窗 1 判定实例（Window 1 checker instance）
    _fbWin2            : FB_DL_TimeWindowCheck;  // 窗 2 判定实例（Window 2 checker instance）
    _fbWin3            : FB_DL_TimeWindowCheck;  // 窗 3 判定实例（Window 3 checker instance）
    _fbWin4            : FB_DL_TimeWindowCheck;  // 窗 4 判定实例（Window 4 checker instance）
    fbTrigReset        : R_TRIG;                 // 复位信号上升沿检测实例（Reset edge detector）
    fbTrigOccupy       : R_TRIG;                 // 占用开始沿检测实例（Occupancy edge detector），CLK = bOccupied
    _eWd               : E_DL_Weekday := E_DL_Weekday.eInvalid;  // 星期换算返回值（Weekday calc result，复用 DL_Base 既有枚举）
    _uErrDow           : UDINT;                  // 星期换算返回码（Weekday calc code）16#0001_0201 = 日期越界
    _bDateOk           : BOOL;                   // 日期有效性（Date valid）
    _uWd               : USINT;                  // 当日星期 USINT 域（Current weekday）1..7，0=非法
    _bWdOk             : BOOL;                   // 星期索引有效性（Weekday index valid）
    _bTimeOk           : BOOL;                   // 当前时刻有效性（Time-of-day valid）
    _abWdSel           : ARRAY[1..7] OF BOOL;    // 单日位展开表（Expanded single-day table），喂窗实例 aWeekdayEnable
    abEnDay            : ARRAY[1..4] OF BOOL;    // 各窗日总使能（Per-window day enable）= 窗使能 AND NOT 节假日覆盖
    abWdBit            : ARRAY[1..4] OF BOOL;    // 各窗当日星期位（Per-window weekday bit）
    abWinValid         : ARRAY[1..4] OF BOOL;    // 各窗今日有效（Per-window valid today）= 日使能 AND 星期位 AND 开启参数合法
    abOccWin           : ARRAY[1..4] OF BOOL;    // 各窗占用结果（Per-window occupancy）
    abPreBand          : ARRAY[1..4] OF BOOL;    // 各窗预启带命中（Per-window pre-start band hit）
    _nNowMin           : DINT;                   // 当前时刻折算分钟（Now in minutes）0..1439，USINT→DINT 扩宽防溢出
    _nStartMin         : DINT;                   // 窗开始折算分钟（Start in minutes）0..1439，扩宽防溢出
    _atStartT          : ARRAY[1..4] OF TIME;    // 各窗开始时刻 TIME 域（Per-window start time），分钟折算防溢出后换域
    _tNowT             : TIME;                   // 当前时刻 TIME 域（Now in TIME domain），预启带比较用
    _tLeadT            : TIME;                   // 生效提前量（Effective lead time）防御钳位 ≤ T#12H
    _i                 : USINT;                  // 循环索引（Loop index）1..4，固定界防死循环
    _j                 : USINT;                  // 循环索引（Loop index）1..7，固定界防死循环
END_VAR

// -----------------------------------------------------------------------------
// 段 1｜复位沿实例无条件周期刷新（R7 红线：严禁移入 IF/CASE 分支）
// -----------------------------------------------------------------------------
fbTrigReset(CLK := bReset);                 // 复位沿检测

// -----------------------------------------------------------------------------
// 段 2｜出口默认值与时刻有效性（事件型逐拍重算，无状态驻留）
// -----------------------------------------------------------------------------
uErrorId := 16#0000_0000;                   // 信息级码每拍重算
bOccupied := FALSE;                         // 占用合成默认 FALSE
bPreStart := FALSE;                         // 预启动默认 FALSE
bPulseOnOccupy := FALSE;                    // 沿单发默认 FALSE（段 10 覆盖）
uActiveWin := 0;                            // 活动窗号默认无
_bTimeOk := (uHourNow <= 23) AND (uMinNow <= 59);   // 时刻域检查（越界预启动跳过）

// -----------------------------------------------------------------------------
// 段 3｜星期换算：FC_DL_DayOfWeekCalc 公开接口直接调用（不内联重实现）
// -----------------------------------------------------------------------------
_eWd := FC_DL_DayOfWeekCalc(uYear := uYear, uMonth := uMonth, uDay := uDay,
                            uErrorId => _uErrDow);              // 日期 → 星期（ISO 序）
_bDateOk := (_uErrDow = 16#0000_0000);                          // 返回码 0 = 日期合法
IF NOT _bDateOk THEN
    uErrorId := 16#0005_0210;               // 日期非法【信息级】：全窗按不在窗处理
END_IF

// 星期枚举 → USINT 索引显式映射（strict 枚举不整型直赋；CASE+ELSE 兜底）
CASE _eWd OF
    E_DL_Weekday.eMonday:    _uWd := 1;     // 周一（ISO 1）
    E_DL_Weekday.eTuesday:   _uWd := 2;     // 周二（ISO 2）
    E_DL_Weekday.eWednesday: _uWd := 3;     // 周三（ISO 3）
    E_DL_Weekday.eThursday:  _uWd := 4;     // 周四（ISO 4）
    E_DL_Weekday.eFriday:    _uWd := 5;     // 周五（ISO 5）
    E_DL_Weekday.eSaturday:  _uWd := 6;     // 周六（ISO 6）
    E_DL_Weekday.eSunday:    _uWd := 7;     // 周日（ISO 7）
    ELSE
        _uWd := 0;                          // eInvalid / 未预期：当日全窗不使能
END_CASE
_bWdOk := (_uWd >= 1) AND (_uWd <= 7);      // 索引域校验（防矩阵越界，R4）

// -----------------------------------------------------------------------------
// 段 4｜公共量预计算：日使能 / 星期位 / 窗有效性 / 开始时刻折算（分钟域扩宽）
// -----------------------------------------------------------------------------
FOR _i := 1 TO 4 DO
    abEnDay[_i] := aWinEnable[_i] AND (NOT aHolidayOverride[_i]);   // 日总使能 = 窗使能 AND NOT 节假日
    abWdBit[_i] := FALSE;                   // 星期位默认 FALSE（索引非法时全窗不使能）
    IF _bWdOk THEN
        abWdBit[_i] := aWeekdayWin[_i, _uWd];   // 当日星期位（索引 1..7 已校验）
    END_IF
    abWinValid[_i] := abEnDay[_i] AND abWdBit[_i]
                   AND (aHourOn[_i] <= 23) AND (aMinOn[_i] <= 59);
                                            // 今日有效 = 日使能 AND 星期位 AND 开启参数合法
    _nStartMin := aHourOn[_i];              // USINT → DINT 扩宽（先赋值再乘防溢出）
    _nStartMin := (_nStartMin * 60) + aMinOn[_i];   // 开窗分钟 0..1439
    _atStartT[_i] := T#1M * _nStartMin;     // 分钟域 → TIME 域（MUL(TIME, 整数) 标准序）
END_FOR

_nNowMin := uHourNow;                       // USINT → DINT 扩宽
_nNowMin := (_nNowMin * 60) + uMinNow;      // 当前分钟 0..1439（越界值仅预启带门控弃用）
_tNowT := T#1M * _nNowMin;                  // 当前时刻 → TIME 域
_tLeadT := tPreLeadTime;                    // 提前量原值生效
IF _tLeadT > T#12H THEN
    _tLeadT := T#12H;                       // 防御钳位：提前量组态域建议 ≤ 半日，回绕式防负时长
END_IF

// -----------------------------------------------------------------------------
// 段 5~8｜窗 1~4 实例逐拍无条件刷新（R7：调用与输入准备均不入 IF/CASE 分支）
//        每窗：单日位展开 → 实例调用 → 占用收集 → 实例码归并 → 预启带判定
// -----------------------------------------------------------------------------

// ---- 窗 1（Window 1）----
FOR _j := 1 TO 7 DO
    _abWdSel[_j] := abWdBit[1];             // aWeekdayWin[1, 当日] 单日位展开为 7 日表
END_FOR
_fbWin1(uHourNow := uHourNow, uMinNow := uMinNow,
        bEnableDay := abEnDay[1], aWeekdayEnable := _abWdSel, uWeekdayNow := _uWd,
        uHourOn := aHourOn[1], uMinOn := aMinOn[1],
        uHourOff := aHourOff[1], uMinOff := aMinOff[1], bReset := FALSE);
                                            // 窗 1 实例刷新（bReset 恒 FALSE：实例码仅当拍归并）
abOccWin[1] := _fbWin1.bInWindow;           // 窗 1 占用结果
IF _bDateOk AND (_fbWin1.uErrorId <> 16#0000_0000) THEN
    uErrorId := 16#0005_0211;               // 实例码不透传，归并为本块 0211【信息级】
END_IF
abPreBand[1] := FALSE;                      // 预启带默认未命中
IF abWinValid[1] AND _bTimeOk THEN
    IF _tLeadT <= _atStartT[1] THEN
        abPreBand[1] := (_tNowT >= (_atStartT[1] - _tLeadT)) AND (_tNowT < _atStartT[1]);
                                            // 同日内预启带 [开始−提前, 开始) 左闭右开
    ELSE
        abPreBand[1] := (_tNowT >= ((_atStartT[1] + T#24H) - _tLeadT))
                    OR (_tNowT < _atStartT[1]);
                                            // 跨零点回绕：预启带 [开始+24h−提前, 24h)∪[0, 开始)
    END_IF
END_IF

// ---- 窗 2（Window 2）----
FOR _j := 1 TO 7 DO
    _abWdSel[_j] := abWdBit[2];             // aWeekdayWin[2, 当日] 单日位展开
END_FOR
_fbWin2(uHourNow := uHourNow, uMinNow := uMinNow,
        bEnableDay := abEnDay[2], aWeekdayEnable := _abWdSel, uWeekdayNow := _uWd,
        uHourOn := aHourOn[2], uMinOn := aMinOn[2],
        uHourOff := aHourOff[2], uMinOff := aMinOff[2], bReset := FALSE);
                                            // 窗 2 实例刷新
abOccWin[2] := _fbWin2.bInWindow;           // 窗 2 占用结果
IF _bDateOk AND (_fbWin2.uErrorId <> 16#0000_0000) THEN
    uErrorId := 16#0005_0211;               // 实例码归并【信息级】
END_IF
abPreBand[2] := FALSE;                      // 预启带默认未命中
IF abWinValid[2] AND _bTimeOk THEN
    IF _tLeadT <= _atStartT[2] THEN
        abPreBand[2] := (_tNowT >= (_atStartT[2] - _tLeadT)) AND (_tNowT < _atStartT[2]);
                                            // 同日内预启带
    ELSE
        abPreBand[2] := (_tNowT >= ((_atStartT[2] + T#24H) - _tLeadT))
                    OR (_tNowT < _atStartT[2]);
                                            // 跨零点回绕预启带
    END_IF
END_IF

// ---- 窗 3（Window 3）----
FOR _j := 1 TO 7 DO
    _abWdSel[_j] := abWdBit[3];             // aWeekdayWin[3, 当日] 单日位展开
END_FOR
_fbWin3(uHourNow := uHourNow, uMinNow := uMinNow,
        bEnableDay := abEnDay[3], aWeekdayEnable := _abWdSel, uWeekdayNow := _uWd,
        uHourOn := aHourOn[3], uMinOn := aMinOn[3],
        uHourOff := aHourOff[3], uMinOff := aMinOff[3], bReset := FALSE);
                                            // 窗 3 实例刷新
abOccWin[3] := _fbWin3.bInWindow;           // 窗 3 占用结果
IF _bDateOk AND (_fbWin3.uErrorId <> 16#0000_0000) THEN
    uErrorId := 16#0005_0211;               // 实例码归并【信息级】
END_IF
abPreBand[3] := FALSE;                      // 预启带默认未命中
IF abWinValid[3] AND _bTimeOk THEN
    IF _tLeadT <= _atStartT[3] THEN
        abPreBand[3] := (_tNowT >= (_atStartT[3] - _tLeadT)) AND (_tNowT < _atStartT[3]);
                                            // 同日内预启带
    ELSE
        abPreBand[3] := (_tNowT >= ((_atStartT[3] + T#24H) - _tLeadT))
                    OR (_tNowT < _atStartT[3]);
                                            // 跨零点回绕预启带
    END_IF
END_IF

// ---- 窗 4（Window 4）----
FOR _j := 1 TO 7 DO
    _abWdSel[_j] := abWdBit[4];             // aWeekdayWin[4, 当日] 单日位展开
END_FOR
_fbWin4(uHourNow := uHourNow, uMinNow := uMinNow,
        bEnableDay := abEnDay[4], aWeekdayEnable := _abWdSel, uWeekdayNow := _uWd,
        uHourOn := aHourOn[4], uMinOn := aMinOn[4],
        uHourOff := aHourOff[4], uMinOff := aMinOff[4], bReset := FALSE);
                                            // 窗 4 实例刷新
abOccWin[4] := _fbWin4.bInWindow;           // 窗 4 占用结果
IF _bDateOk AND (_fbWin4.uErrorId <> 16#0000_0000) THEN
    uErrorId := 16#0005_0211;               // 实例码归并【信息级】
END_IF
abPreBand[4] := FALSE;                      // 预启带默认未命中
IF abWinValid[4] AND _bTimeOk THEN
    IF _tLeadT <= _atStartT[4] THEN
        abPreBand[4] := (_tNowT >= (_atStartT[4] - _tLeadT)) AND (_tNowT < _atStartT[4]);
                                            // 同日内预启带
    ELSE
        abPreBand[4] := (_tNowT >= ((_atStartT[4] + T#24H) - _tLeadT))
                    OR (_tNowT < _atStartT[4]);
                                            // 跨零点回绕预启带
    END_IF
END_IF

// -----------------------------------------------------------------------------
// 段 9｜占用合成与活动窗号（多窗同开取最小号；日期非法时全窗自然为 FALSE）
// -----------------------------------------------------------------------------
bOccupied := abOccWin[1] OR abOccWin[2] OR abOccWin[3] OR abOccWin[4];
                                            // 任一有效窗在窗内即占用
FOR _i := 1 TO 4 DO
    IF abOccWin[_i] AND (uActiveWin = 0) THEN
        uActiveWin := _i;                   // 取最小活动窗号（升序首中）
    END_IF
END_FOR

bPreStart := (NOT bOccupied) AND _bTimeOk
         AND (abPreBand[1] OR abPreBand[2] OR abPreBand[3] OR abPreBand[4]);
                                            // 预启动：未占用 AND 时刻合法 AND 任一有效窗预启带命中

// -----------------------------------------------------------------------------
// 段 10｜占用开始沿单发（实例无条件周期刷新，沿输出持续一拍）
// -----------------------------------------------------------------------------
fbTrigOccupy(CLK := bOccupied);             // 占用上升沿检测（主体无条件调用）
bPulseOnOccupy := fbTrigOccupy.Q;           // 占用开始沿单发输出

// -----------------------------------------------------------------------------
// 段 11｜复位沿消费：清除当拍信息级码（触发实例已在段 1 无条件刷新）
// -----------------------------------------------------------------------------
IF fbTrigReset.Q THEN
    uErrorId := 16#0000_0000;               // 复位沿当拍清信息级码（下一拍重新评估）
END_IF

END_FUNCTION_BLOCK

(* ---- FB_DL_PalletizerLayerBuildSeq.st ---- *)
(*==============================================================================
 * 组件名称 (Component)  : FB_DL_PalletizerLayerBuildSeq
 * 所属子库 (Sublibrary) : DL_Process ｜ 版本 (Version) : 1.0.2 ｜ 2026-11-23
 * 兼容性   (Platform)   : CODESYS 3.5+ / TwinCAT 3 / 汇川 InoProShop / 施耐德 Machine Expert
 *                         仅依赖 IEC 61131-3 标准库（TON 属 Standard.library），零厂商私有库
 * 功能描述 (Function)   : 码垛层构建时序：eIdle →（bStart）→ ePick（发取料指令，等
 *                         bPickDone 到位）→ ePlace（发放料指令，等 bPlaceDone 到位并计数）
 *                         → 满层判（nPlacedInLayer ≥ nBoxPerLayer）→ eLayerDone（发单拍层完成沿）
 *                         → 换层（nLayerNo + 1，层内计数清零）回 ePick；层数达 nLayersPerPallet
 *                         → eFull（整垛完成，等 bStart 跌落或复位）。取 / 放每相均带
 *                         tPhaseTimeout 超时兜底 → eFault。
 *                         **输出语义**：bPickCmd / bPlaceCmd 为电平台（相驻留期间为 TRUE），
 *                         bLayerDone 为**单拍脉冲**（内部 _bLayerDoneInt 置位 → 统一出口映射，
 *                         两段式，FB33-1），每拍由段 1 预置 FALSE，故脉冲宽度恰一扫描。
 *                         **bStart = FALSE 语义（R191 二选一，本件选「降级为安全值 + 置标志」）**：
 *                         全部动作输出落 FALSE 并回 eIdle（码垛动作不得冻结保持，冻结即撞机）。
 * 接口     (Interface)  : 输入 bStart / bReset / bPickDone / bPlaceDone / nBoxPerLayer /
 *                         nLayersPerPallet / tPhaseTimeout；输出 bPickCmd / bPlaceCmd /
 *                         nPlacedInLayer / nLayerNo / bLayerDone / bPalletFull / eState /
 *                         bError / eCause / bValid。
 * 状态迁移表 (State Transition Table)：
 *   ① eIdle → ePick：bStart 为 TRUE 且组态校验通过（nBoxPerLayer / nLayersPerPallet 均在域内）；
 *      拍 N 进入（启动）/ 本拍行为：层内计数与层号初始化（nPlacedInLayer := 0、nLayerNo := 1）、
 *      不发指令 / 拍 N+1 转出至 ePick。
 *   ② ePick → ePlace：bPickDone 上升沿（本拍事件优先于超时，FB51-5）；拍 N 进入（取料到位）/
 *      本拍行为：撤 bPickCmd、发 bPlaceCmd / 拍 N+1 转出至 ePlace。
 *   ③ ePick → eFault：tonPhase.Q（超时）；拍 N 进入（超时）/ 本拍行为：锁存 ePickTimeout、
 *      撤全部动作 / 拍 N+1 转出至 eFault（段尾迁移闸）。
 *   ④ ePlace → ePick：bPlaceDone 上升沿且层未满（nPlacedInLayer + 1 < nBoxPerLayer）；
 *      拍 N 进入（放料到位）/ 本拍行为：层内计数 +1、撤 bPlaceCmd / 拍 N+1 转出至 ePick。
 *   ⑤ ePlace → eLayerDone：bPlaceDone 上升沿且本次计数后层已满；拍 N 进入 /
 *      本拍行为：层内计数 +1、_bLayerDoneInt := TRUE / 拍 N+1 转出至 eLayerDone。
 *   ⑥ ePlace → eFault：tonPhase.Q（超时），锁存 ePlaceTimeout。
 *   ⑦ eLayerDone → eFull：nLayerNo ≥ nLayersPerPallet；拍 N 进入 / 本拍行为：bPalletFull := TRUE /
 *      拍 N+1 转出至 eFull。
 *   ⑧ eLayerDone → ePick：层未满垛；拍 N 进入 / 本拍行为：nLayerNo + 1、nPlacedInLayer := 0 /
 *      拍 N+1 转出至 ePick。
 *   ⑨ eFull → eIdle：bStart 落 FALSE（前置条件消失）或 bReset 为 TRUE（两条出口，R98）；
 *      拍 N 进入 / 本拍行为：层号与层内计数清零、bPalletFull 落 FALSE / 拍 N+1 转出至 eIdle。
 *   ⑩ eFault → eIdle：bReset 上升且 bStart 为 FALSE（可达性自证 R152：两引脚外部恒可达）；
 *      拍 N 进入 / 本拍行为：清锁存与成因 / 拍 N+1 转出至 eIdle。
 *   ⑪ ELSE（非法枚举值）→ eFault，成因 eIllegalState（R6 兜底）。
 * 边界     (Boundary)   : ① 相超时 TON 在 CASE 外无条件调用（R7 / FB50-1①），IN 表达式为
 *                            「处于取/放相 AND 相已稳定一拍（nPhase = nPhasePrev）AND
 *                            非故障相 AND 非故障锁存」——相切换那一拍 IN 为 FALSE 使 ET 自清，
 *                            结构性无需外部沿清零（R188）。
 *                         ② 组态域闸：nBoxPerLayer ∈ [1,60]、nLayersPerPallet ∈ [1,40]，
 *                            越域置故障级 eBadConfig（R4，兼作数组/计数安全）。
 *                         ③ ePick / ePlace 退出条件均为「事件沿 + 超时」两条（R98）。
 *                         ④ 无数组、无除法，故无下标与除零风险。
 *                         ⑤ 零全局耦合（无 GVL / VAR_EXTERNAL / %I / %Q）。
 * 码表     (Codes)      : 本件不占用全局数字码位（R297 零码位范式）；出口为 BOOL + ENUM，
 *                         enum E_DL_PlbCause 归属本文件（全库唯一属主）。信息级
 *                         eLayerDoneCode 永不置 bError；超时 / 组态 / 非法状态各占独立成员
 *                         （R190 归因唯一），锁存回放至 bReset 沿（FB33-1）。
 * 分工声明 (Scope)      : 层内路径规划 / 码型排布归 FB_DL_PalletizerStation 与
 *                         FB_DL_PalletizerLayerSeq（区段时序）；夹爪安全归 FB_DL_PalletGripperSafe。
 *                         本件只做「取—放—满层—换层—满垛」的计数与时序，不做轴运动与轨迹。
 * 归属     (Ownership)  : E_DL_PlbState / E_DL_PlbCause 归属本文件（全库唯一定义，R264）。
 * 红线自检 (Redline)    : R1 ✓ 零 GVL ｜ R2 ✓ 零 %I/%Q ｜ R3 ✓ 纯 IEC ｜ R4 ✓ 组态域闸 +
 *                         无除法无下标 + 计数单调 ｜ R5 ✓ 逐行同行双语注释 ｜ R6 ✓ 六态 ENUM +
 *                         CASE + ELSE ｜ R7 ✓ tonPhase 在 CASE 外无条件调用 ｜ R14 ✓ 无 PROPERTY
 *                         R8/R9 N/A（无 METHOD）｜ FB32-6 ✓ 单拍脉冲置位与撤销分属两拍
 * 修订历史 (Revision)   : 2026-11-23  v1.0.0  R78-B3 首版
 * 验收向量 (Acceptance) :
 *   V1 nBoxPerLayer=2、nLayersPerPallet=2：bStart 上升 → ePick；bPickDone 脉冲 → ePlace；
 *      bPlaceDone 脉冲 → nPlacedInLayer=1 且回 ePick；再一轮 → nPlacedInLayer=2、eLayerDone、
 *      bLayerDone 单拍为 TRUE（次拍 FALSE）；随后 nLayerNo=2、nPlacedInLayer=0、ePick。
 *   V2 续 V1 完成第 2 层 → eFull、bPalletFull=TRUE；bStart 落 FALSE → 回 eIdle，计数全清。
 *   V3 tPhaseTimeout=5s、bPickDone 始终不来 → 5s 后 eState=eFault、eCause=ePickTimeout、
 *      bError=TRUE、bPickCmd=FALSE；bReset 上升且 bStart=FALSE → 回 eIdle。
 *   V4 nBoxPerLayer=0 → eState=eFault、eCause=eBadConfig、bError=TRUE。
 *   V5 eFull 内 bReset=TRUE（bStart 仍 TRUE）→ 回 eIdle 并清计数（第二条出口）。
 *============================================================================*)

(*-----------------------------------------------------------------------------
 * 枚举: E_DL_PlbState（码垛层构建相位；eFault 为安全相，仅 bReset 沿迁出）
 *----------------------------------------------------------------------------*)
TYPE E_DL_PlbState :
(
    eIdle      := 0,    // 空闲：无动作输出，等 bStart / Idle: no motion command, waiting for bStart
    ePick      := 10,   // 取料相：bPickCmd 电平为 TRUE，等 bPickDone / Pick phase: bPickCmd high until bPickDone
    ePlace     := 20,   // 放料相：bPlaceCmd 电平为 TRUE，等 bPlaceDone / Place phase: bPlaceCmd high until bPlaceDone
    eLayerDone := 30,   // 层完成相：发 bLayerDone 单拍沿并判定换层 / Layer done: emit the single-scan edge and decide
    eFull      := 40,   // 整垛完成相：bPalletFull 电平为 TRUE / Pallet full: bPalletFull high
    eFault     := 90    // 故障安全相：超时 / 组态非法，动作全撤 / Fault safe phase: timeout or bad configuration
);
END_TYPE

(*-----------------------------------------------------------------------------
 * 枚举: E_DL_PlbCause（成因码；信息级 = 0..9，故障级 = 10 起）
 *----------------------------------------------------------------------------*)
TYPE E_DL_PlbCause :
(
    eNone          := 0,   // 信息级：无事件 / Info: no event
    eLayerDoneCode := 1,   // 信息级：一层已构建完成 / Info: one layer completed
    ePalletDone    := 2,   // 信息级：整垛完成 / Info: pallet completed
    ePickTimeout   := 10,  // 故障级：取料相超时 / Fault: pick phase timeout
    ePlaceTimeout  := 11,  // 故障级：放料相超时 / Fault: place phase timeout
    eBadConfig     := 12,  // 故障级：每层箱数 / 每垛层数越域 / Fault: box-per-layer or layer count out of domain
    eIllegalState  := 13   // 故障级：非法状态枚举值 / Fault: illegal state enum value
);
END_TYPE

FUNCTION_BLOCK FB_DL_PalletizerLayerBuildSeq
VAR_INPUT
    bStart          : BOOL := FALSE;          // 启动（电平）：FALSE 时动作全撤并回 eIdle / Start level, FALSE withdraws all commands
    bReset          : BOOL := FALSE;          // 复位（上升沿，需同时 bStart=FALSE）/ Reset rising edge, requires bStart FALSE
    bPickDone       : BOOL := FALSE;         // 取料到位反馈（上升沿表示本相完成，初值 FALSE 防首拍假沿）/ Pick completion feedback, rising edge ends the phase, FALSE default avoids a first-scan ghost edge
    bPlaceDone      : BOOL := FALSE;         // 放料到位反馈（上升沿表示本相完成，初值 FALSE 防首拍假沿）/ Place completion feedback, rising edge ends the phase, FALSE default avoids a first-scan ghost edge
    nBoxPerLayer    : INT := 5;               // 每层箱数，有效域 1..60 [-] / Boxes per layer, valid domain 1..60
    nLayersPerPallet : INT := 6;              // 每垛层数，有效域 1..40 [-] / Layers per pallet, valid domain 1..40
    tPhaseTimeout   : TIME := T#10S;          // 单相超时（取/放共用），域 > 0 [s] / Phase timeout shared by pick and place
END_VAR
VAR_OUTPUT
    bPickCmd        : BOOL;                   // 取料指令（电平）/ Pick command, level signal
    bPlaceCmd       : BOOL;                   // 放料指令（电平）/ Place command, level signal
    nPlacedInLayer  : INT := 0;               // 本层已放箱数 [个] / Boxes placed in the current layer
    nLayerNo        : INT := 0;               // 当前层号（1 起）[层] / Current layer number starting at one
    bLayerDone      : BOOL;                   // 层完成单拍脉冲（段 1 预置，统一出口映射）[-] / Single-scan layer-done pulse
    bPalletFull     : BOOL;                   // 整垛完成（电平，保持至 bStart 跌落或复位）[-] / Pallet full, level held until bStart falls or reset
    eState          : E_DL_PlbState;           // 状态出口（段尾单点映射）[-] / State outlet mapped at the tail
    bError          : BOOL;                   // 故障锁存标志 [-] / Fault latch flag
    eCause          : E_DL_PlbCause;          // 成因码出口（故障期锁存回放）[-] / Cause code outlet
    bValid          : BOOL;                   // 时序有效回执（取/放相才 TRUE）[-] / Sequence validity receipt
END_VAR
VAR
    _eState        : E_DL_PlbState := E_DL_PlbState.eIdle;    // 内部相位（CASE 唯一写入目标）[-] / Internal phase
    _eStatePrev    : E_DL_PlbState := E_DL_PlbState.eIdle;    // 上一拍相位快照（相稳定判据用，段末唯一更新）[-] / Phase snapshot of the last scan
    _bFaultLatch   : BOOL := FALSE;                           // 故障锁存位（仅 bReset 沿清除）[-] / Fault latch bit
    _eCauseLatch   : E_DL_PlbCause := E_DL_PlbCause.eNone;     // 锁存成因码（FB33-1 锁存回放）[-] / Latched cause code
    _bCfgOk        : BOOL := TRUE;                            // 组态域闸通过标志 [-] / Configuration gate flag
    _bLayerDoneInt : BOOL := FALSE;                           // 层完成内部单拍位（统一出口映射，FB33-1）[-] / Internal single-scan layer-done bit
    _bPhaseActive  : BOOL := FALSE;                           // 取/放相驻留标志（超时使能域）[-] / Phase-resident flag driving the timeout
    _bPickRise     : BOOL := FALSE;                           // 取料到位上升沿（本拍）/ Pick completion rising edge of this scan
    _bPlaceRise    : BOOL := FALSE;                           // 放料到位上升沿（本拍）/ Place completion rising edge of this scan
    rtPickDone     : R_TRIG;                                  // 取料到位边沿实例（段 3 无条件调用）/ Pick edge instance called unconditionally
    rtPlaceDone    : R_TRIG;                                  // 放料到位边沿实例（段 3 无条件调用）/ Place edge instance called unconditionally
    tonPhase       : TON;                                     // 相超时定时器（段 3 无条件调用）/ Phase timeout timer called unconditionally
    _rtReset     : R_TRIG;                                 // 复位沿检测实例（v1.0.2 补：声明沿即实现沿，CASE 外无条件刷新）/ Reset edge detector refreshed outside the CASE
END_VAR
VAR CONSTANT
    DL_PLB_ZERO      : INT := 0;      // 计数零基准 [-] / Count zero base
    DL_PLB_ONE       : INT := 1;      // 计数起始值（层号与每层首箱）[-] / Count start value
    DL_PLB_BOX_MAX   : INT := 60;     // 每层箱数上限（域闸用）[-] / Upper bound of boxes per layer
    DL_PLB_LAYER_MAX : INT := 40;     // 每垛层数上限（域闸用）[-] / Upper bound of layers per pallet
END_VAR

(* —— 段 1：单拍位与动作出口预置（纸清单拍标志与电平出口，不清锁存/计数，FB32-1） —— *)
bLayerDone     := FALSE;                                // 单拍层完成沿每拍预清 / Single-scan edge preset FALSE every scan
bPickCmd       := FALSE;                                // 取料指令预置（安全侧：默认不动作）/ Pick command preset, safe side
bPlaceCmd      := FALSE;                                // 放料指令预置（安全侧：默认不动作）/ Place command preset, safe side
_bLayerDoneInt := FALSE;                                // 内部单拍位预清 / Internal single-scan bit preset
_bCfgOk        := TRUE;                                 // 组态闸标志复位 / Configuration flag reset

(* —— 段 2：组态域闸（每层箱数 / 每垛层数，R4） —— *)
IF (nBoxPerLayer < DL_PLB_ONE) OR (nBoxPerLayer > DL_PLB_BOX_MAX)
    OR (nLayersPerPallet < DL_PLB_ONE) OR (nLayersPerPallet > DL_PLB_LAYER_MAX) THEN
    _bCfgOk := FALSE;                                   // 组态越域 / Configuration out of domain
    IF NOT _bFaultLatch THEN
        _eCauseLatch := E_DL_PlbCause.eBadConfig;       // 故障级：组态非法（首因锁存）/ Fault: bad configuration
        _bFaultLatch := TRUE;                           // 置故障锁存 / Latch the fault
    END_IF
END_IF

(* —— 段 3：边沿与超时实例（CASE 外无条件调用，R7 / FB50-1①） —— *)
rtPickDone(CLK := bPickDone);                           // 取料到位沿（无条件刷新：非取料相期间的沿被吞，属 R7 固有口径）/ Pick completion edge, refreshed unconditionally, edges outside the phase are consumed
rtPlaceDone(CLK := bPlaceDone);                         // 放料到位沿（无条件刷新，沿吞噬口径与取料沿一致）/ Place completion edge, refreshed unconditionally with the same edge-consumption rule
_bPickRise  := rtPickDone.Q;                            // 取料沿快照 / Pick edge snapshot
_bPlaceRise := rtPlaceDone.Q;                           // 放料沿快照 / Place edge snapshot
_bPhaseActive := (_eState = E_DL_PlbState.ePick) OR (_eState = E_DL_PlbState.ePlace);   // 取/放相驻留 / Phase residency
tonPhase(IN := _bPhaseActive AND (_eState = _eStatePrev) AND (_eState <> E_DL_PlbState.eFault) AND (NOT _bFaultLatch),
         PT := tPhaseTimeout);                          // 相稳定一拍后才计时，相切换拍 ET 自清（R188）/ Timer armed only after a stable phase scan

(* —— 段 4：状态机主体（唯一相位写入点，事件沿优先于超时，FB51-5） —— *)
_rtReset(CLK := bReset);                                // 复位沿刷新无条件周期调用（R7；v1.0.2 修复 J1 电平判据缺陷 / R18）/ Refresh the reset edge unconditionally every scan
CASE _eState OF
    E_DL_PlbState.eIdle :
        IF bStart AND (NOT _bFaultLatch) THEN
            nPlacedInLayer := DL_PLB_ZERO;              // 层内计数清零 / Clear the in-layer count
            nLayerNo       := DL_PLB_ONE;               // 层号置 1 / Start at layer one
            bPalletFull    := FALSE;                    // 整垛标志复位 / Clear the pallet-full flag
            eCause         := E_DL_PlbCause.eNone;      // 信息级：无事件 / Info: no event
            _eState        := E_DL_PlbState.ePick;      // 迁移①：进入取料相 / Move to pick
        ELSE
            bPalletFull := FALSE;                       // 未启动：整垛标志保持 FALSE / Not started: pallet flag FALSE
        END_IF

    E_DL_PlbState.ePick :
        bPickCmd := TRUE;                               // 取料指令电平为 TRUE / Pick command high
        IF _bPickRise THEN
            (* 迁移②：本拍事件优先，先消化到位沿再消化超时（FB51-5） *)
            bPickCmd := FALSE;                          // 撤取料指令 / Withdraw the pick command
            eCause   := E_DL_PlbCause.eNone;            // 信息级：无事件 / Info: no event
            _eState  := E_DL_PlbState.ePlace;           // 迁入放料相 / Move to place
        ELSIF tonPhase.Q THEN
            (* 迁移③：超时兜底 *)
            _eCauseLatch := E_DL_PlbCause.ePickTimeout; // 故障级：取料超时 / Fault: pick timeout
            _bFaultLatch := TRUE;                       // 置故障锁存 / Latch the fault
            bPickCmd     := FALSE;                      // 撤动作 / Withdraw the command
            _eState      := E_DL_PlbState.eFault;       // 迁入故障相 / Move to fault
        END_IF

    E_DL_PlbState.ePlace :
        bPlaceCmd := TRUE;                              // 放料指令电平为 TRUE / Place command high
        IF _bPlaceRise THEN
            (* 迁移④ / ⑤：放料到位 → 计数 + 满层判（两出口分列） *)
            bPlaceCmd      := FALSE;                    // 撤放料指令 / Withdraw the place command
            nPlacedInLayer := nPlacedInLayer + DL_PLB_ONE;   // 层内计数 +1 / Increment the in-layer count
            IF nPlacedInLayer >= nBoxPerLayer THEN
                _bLayerDoneInt := TRUE;                 // 层已满：内部单拍位置位（统一出口映射）/ Layer full: internal edge bit
                eCause         := E_DL_PlbCause.eLayerDoneCode;   // 信息级：一层完成 / Info: one layer done
                _eState        := E_DL_PlbState.eLayerDone;       // 迁入层完成相 / Move to layer done
            ELSE
                eCause := E_DL_PlbCause.eNone;          // 信息级：无事件 / Info: no event
                _eState := E_DL_PlbState.ePick;         // 回取料相继续本层 / Back to pick for the same layer
            END_IF
        ELSIF tonPhase.Q THEN
            (* 迁移⑥：超时兜底 *)
            _eCauseLatch := E_DL_PlbCause.ePlaceTimeout;   // 故障级：放料超时 / Fault: place timeout
            _bFaultLatch := TRUE;                          // 置故障锁存 / Latch the fault
            bPlaceCmd    := FALSE;                         // 撤动作 / Withdraw the command
            _eState      := E_DL_PlbState.eFault;          // 迁入故障相 / Move to fault
        END_IF

    E_DL_PlbState.eLayerDone :
        IF nLayerNo >= nLayersPerPallet THEN
            bPalletFull := TRUE;                        // 迁移⑦：整垛满 / Pallet full
            eCause      := E_DL_PlbCause.ePalletDone;   // 信息级：整垛完成 / Info: pallet completed
            _eState     := E_DL_PlbState.eFull;         // 迁入整垛完成相 / Move to full
        ELSE
            nLayerNo       := nLayerNo + DL_PLB_ONE;    // 迁移⑧：换层 / Next layer
            nPlacedInLayer := DL_PLB_ZERO;              // 层内计数清零 / Clear the in-layer count
            eCause         := E_DL_PlbCause.eNone;      // 信息级：无事件 / Info: no event
            _eState        := E_DL_PlbState.ePick;      // 回取料相 / Back to pick
        END_IF

    E_DL_PlbState.eFull :
        (* 迁移⑨：两条出口（前置条件消失 / 复位），R98 *)
        IF (NOT bStart) OR bReset THEN
            bPalletFull    := FALSE;                    // 整垛标志撤销 / Withdraw the pallet flag
            nPlacedInLayer := DL_PLB_ZERO;              // 层内计数清零 / Clear the in-layer count
            nLayerNo       := DL_PLB_ZERO;              // 层号清零 / Clear the layer number
            eCause         := E_DL_PlbCause.eNone;      // 信息级：无事件 / Info: no event
            _eState        := E_DL_PlbState.eIdle;      // 回空闲相 / Back to idle
        END_IF

    E_DL_PlbState.eFault :
        (* 迁移⑩：唯一出口 —— bReset 沿 + bStart 已落 *)
        IF _rtReset.Q AND (NOT bStart) THEN
            _bFaultLatch   := FALSE;                    // 清故障锁存 / Clear the latch
            _eCauseLatch   := E_DL_PlbCause.eNone;      // 清锁存成因 / Clear the latched cause
            eCause         := E_DL_PlbCause.eNone;      // 出口同步归零 / Outlet follows
            nPlacedInLayer := DL_PLB_ZERO;              // 计数清零 / Clear the count
            nLayerNo       := DL_PLB_ZERO;              // 层号清零 / Clear the layer number
            _eState        := E_DL_PlbState.eIdle;      // 回空闲相 / Back to idle
        END_IF

ELSE
    (* 迁移⑪：非法枚举兜底（R6） *)
    _eCauseLatch := E_DL_PlbCause.eIllegalState;        // 故障级：非法状态 / Fault: illegal state
    _bFaultLatch := TRUE;                               // 置锁存 / Latch
    _eState      := E_DL_PlbState.eFault;               // 迁入故障相 / Move to fault
END_CASE

(* —— 段 5：段尾故障迁移闸（锁存与迁相分离，FB50-1④），动作输出在故障相全撤 —— *)
IF _bFaultLatch AND (_eState <> E_DL_PlbState.eFault) THEN
    _eState := E_DL_PlbState.eFault;                    // 锁存即迁相 / Latch forces the fault phase
END_IF
IF _eState = E_DL_PlbState.eFault THEN
    bPickCmd  := FALSE;                                 // 故障相撤取料 / Fault phase: withdraw pick
    bPlaceCmd := FALSE;                                 // 故障相撤放料 / Fault phase: withdraw place
END_IF

(* —— 段 6：统一出口（状态映射 + 单拍位映射 + 锁存回放） —— *)
eState     := _eState;                                  // 相位映射 / Phase mapping
bLayerDone := _bLayerDoneInt;                           // 单拍层完成沿统一映射（FB33-1 两段式）/ Single-scan edge mapped here
bError     := _bFaultLatch;                             // 故障标志取锁存位 / Fault flag from the latch
IF _bFaultLatch THEN
    eCause := _eCauseLatch;                             // 故障期回放锁存码 / Replay the latched code
END_IF
bValid := _bPhaseActive AND (NOT _bFaultLatch);         // 仅取/放相且无锁存时有效 / Valid only in pick or place without a latch
_eStatePrev := _eState;                                 // 相位快照更新（唯一写入点，超时相稳定判据用）/ Phase snapshot update, single write point
END_FUNCTION_BLOCK

(* ---- FB_DL_PickAndPlaceStation.st ---- *)
(*==============================================================================
 * 组件名称 (Component)  : FB_DL_PickAndPlaceStation
 * 所属子库 (Sublibrary) : DL_Process
 * 当前版本 (Version)    : 1.0.1
 * 组件分类 (Category)   : 功能块（FUNCTION_BLOCK）· 工站模板 · 九步序
 * 兼容性   (Platform)   : CODESYS 3.5 / TwinCAT 3 / 汇川 InoProShop / Schneider
 *                         Machine Expert；仅 Standard.library 的 TON / R_TRIG，
 *                         轴与真空一律经既有接口引用注入，块内零硬件细节
 * 功能描述 (Function)   : 标准「取 升 移 放」上下料工站模板：注入三轴（X/Y/Z）
 *                         与真空发生器接口，按九步序执行单件搬运（确认原点、
 *                         移到取料位、下降、吸取确认、抬升、横移、下降、破真空、
 *                         抬升回原点），含真空建立超时、就位确认、节拍统计与
 *                         安灯级联出口。
 * 状态机规模 (Scope)    : 本块只做工站内工序的七态最小子集（待机、启动自检、
 *                         执行、保持中、已保持、中止收尾、故障）。完整的十七态
 *                         包装机状态机由 FB_DL_PackMlStateMachine 承载，本块
 *                         不重复实现，避免两套全状态机在同一工站内打架。
 * 接口适配说明 (Adapter) : 既有 I_DL_MotionAxis 的属性集不含「到位布尔位」，
 *                         故每步的到位判据写死为「轴处于待机态且位置落在容差
 *                         窗口内」，等价于驱动层的到位位，且不依赖任何厂商
 *                         专用属性；真空侧的吸取与破真空分别映射到既有
 *                         CmdEvacuate 与 CmdBlowOff，方法名与本块语义一一对应。
 * 时间口径 (Time base)  : 节拍以整循环超时定时器的已历时值作秒表，经
 *                         TIME_TO_DINT 转毫秒整数入滑动窗口；该转换族在三个
 *                         主流平台均提供但不属 IEC 61131-3 基础转换表，故此处
 *                         显式声明依赖，若目标平台缺失请改用显式类型转换语法，
 *                         禁止用 TIME 直接除以整数（后者跨平台必错）。
 * 设计要点 (Key notes)  : ① 单步三段式：下发（只发一次）→ 等条件 → 单拍推进，
 *                           动作指令绝不每拍重发；
 *                         ② 步超时统一由一个定时器监视，进入故障前把步号映射为
 *                           对应故障码，现场据此一步定位；
 *                         ③ 缺料与放料位占用属业务态：置安灯与信息级码，不锁
 *                           故障，产线可继续等待上料；
 *                         ④ 真空未建立属本件 NG：计数加一、置安灯、回步一，
 *                           不锁故障（吸盘老化是常态，停线代价更大）；
 *                         ⑤ 搬运中掉件属故障：立即中止并把工件当作已损坏，
 *                           转中止收尾（抬 Z、破真空），避免二次撞机；
 *                         ⑥ 保持态不重发任何运动指令，释放后从当前步继续，
 *                           已完成步不重做。
 * 开源溯源 (Origin)     : packml-omac / tcopen-component。参考 PackML 与 OMAC
 *                         公开的工站级状态语义（只在可执行子集内取七态）与
 *                         TcOpen 公开组件库的契约实现分离、状态只读属性思想。
 *                         仅借状态命名与分层思想，九步序、码位与实现 100% 自有
 *                         clean-room，不构成衍生作品。
 * 依赖     (Depends)    : I_DL_MotionAxis（DL_Motion）、I_DL_VacuumGenerator
 *                         （DL_Device），均为已入库接口，本块不依赖本轮任何新件
 * 故障码表 (Error codes):
 *   16#0005_01B0【信息级】Z 轴原点未就绪超时（保持本步重试）
 *   16#0005_01B1【信息级】真空未建立，本件判 NG
 *   16#0005_01B2【信息级】前置条件不满足（缺料或放料位占用），业务态加安灯
 *   16#0005_01B3【信息级】正常中止完成
 *   16#0005_01B4【信息级】节拍统计窗重建
 *   16#0005_02B0【故障级】X 轴取料位超时
 *   16#0005_02B1【故障级】Z 轴下降取料超时
 *   16#0005_02B2【故障级】Z 轴抬升超时
 *   16#0005_02B3【故障级】X 轴横移超时
 *   16#0005_02B4【故障级】搬运中掉件
 *   16#0005_02B5【故障级】破真空超时
 *   16#0005_02B6【故障级】回原点超时
 *   16#0005_02B7【故障级】非法状态或非法步号兜底
 * 验收向量 (Acceptance) :
 *   V1 正常单件：前置满足、启动一拍 → 步 1 到 9 推进，完成脉冲单拍、
 *      合格计数 1、节拍大于 0、回待机
 *   V2 缺料：在位信号为假即启动 → 停待机、安灯为真、码 01B2、不锁故障
 *   V3 真空失败：步 4 真空确认恒假且吸附计时到 → 不合格计数 1、安灯为真、
 *      回步 1、不锁故障
 *   V4 掉件：步 7 真空确认丢失 → 掉件标志为真、码 02B4、转中止并抬 Z
 *   V5 保持恢复：步 5 完成时给保持 → 进已保持态；释放后从步 6 继续
 *   V6 超时：步 6 长期不到位、单步超时 1 秒 → 码 02B3、进故障、轴停止被调一次
 *   V7 节拍平均：连做 9 件 → 平均节拍只反映最近 8 件
 * 红线自检 (Redline)    : R1 零全局变量表与外部变量引用 ｜ R2 零物理地址直写
 *                         R3 纯 IEC 61131-3 加既有接口 ｜ R4 到位判定用容差、
 *                         接口引用先判有效性、数组索引经模运算保证在窗内
 *                         R5 全变量中英双语同行注释 ｜ R6 ENUM 加 CASE 加 ELSE 兜底
 *                         R7 四个 TON 与两个 R_TRIG 全部在 CASE 之外无条件刷新
 * 修订历史 (Revision)   :
 *   2026-11-15  v1.0.0  首版入库（Round 10 · ROADMAP 工站模板补齐）
 *   2026-11-15  v1.0.1  R10 终审修复三处（均为机检盲区，逐拍推演发现）：
 *                       R-FIX-1【致命】主状态机 CASE 缺 eExecute 标签，执行态
 *                       落入 ELSE 兜底被判非法状态并锁故障，工站永不执行；
 *                       R-FIX-2【严重】进故障时对四路接口一律判空后再调用，
 *                       原实现对未注入的可选 Y 轴直接调用 Stop，属空引用调用；
 *                       R-FIX-3【中等】步 1 下发分支删除 uErrorId 清零语句，
 *                       原写法把同拍刚置位的 01B0 立即覆盖，诊断不可见。
 * 规格偏离登记 (Deviations):
 *   D1 新增 fSafeZ（安全抬升位）与 fPosTol（到位容差）两个输入引脚：规格书
 *      仅以「安全位」文字描述抬升目标、以「到位」文字描述判据，未给引脚；
 *      按八、无魔法数红线提为引脚，向后兼容（有默认值），不改变既有引脚语义。
 *   D2 到位判据不引用 I_DL_MotionAxis 的到位位（该接口无此属性），改为
 *      「eState = eStandstill 且位置落在容差窗内」，等价语义，已写入头注释。
 *   D3 整循环超时沿用 02B7（非法状态兜底码）：本组件码位块 01B0~01B4 与
 *      02B0~02B7 已全部占用，按 R30「不得跨块取号」不得新增 02B8，故复用
 *      兜底码并在注释写明「循环超时同样按兜底处理」，待下一 MAJOR 拆分码位。
 *============================================================================*)

(*------------------------------------------------------------------------------
 * 枚举: E_DL_SpState（唯一主状态机枚举，同名供输出对外可观测，禁止再设第二套）
 *-----------------------------------------------------------------------------*)
TYPE E_DL_SpState :
(
    eIdle     := 0,     // 待机：未启动 / Idle, not started
    eStarting := 5,     // 启动自检：轴就绪、原点就绪、放料位空闲、取料位有件 / Starting self-check
    eExecute  := 10,    // 执行：九步序推进 / Execute, running the nine-step sequence
    eHolding  := 20,    // 保持中：单拍过渡态 / Holding, a single-cycle transition state
    eHeld     := 25,    // 已保持：不重发任何运动指令 / Held, no motion command is re-issued
    eAborting := 30,    // 中止收尾：抬 Z 与破真空，逐拍推进 / Aborting, one command per cycle
    eFault    := 99     // 故障锁定：仅复位沿可退 / Fault latched, only a reset edge leaves
);
END_TYPE

FUNCTION_BLOCK FB_DL_PickAndPlaceStation
VAR_INPUT
    bEnable       : BOOL := TRUE;      // 工站使能 [-] / Station enable
    bStart        : BOOL;              // 启动单件循环，上升沿，已保持态下无效 [-] / Start one cycle on a rising edge, ignored while held
    bHold         : BOOL;              // 保持，电平：当前步完成后停在已保持态 [-] / Hold, level: park after the current step completes
    bAbort        : BOOL;              // 中止，电平：任何态转中止收尾 [-] / Abort, level: any state goes to the abort sequence
    bReset        : BOOL;              // 复位故障，上升沿 [-] / Reset the fault on a rising edge
    bPartPresent  : BOOL;              // 取料位工件在位（光电）[-] / Part present at the pick position
    bPlaceClear   : BOOL;              // 放料位空闲，允许放料 [-] / Place position clear
    bVacuumOk     : BOOL;              // 真空建立确认（真空开关）[-] / Vacuum established confirmation
    bZHomeOk      : BOOL;              // Z 轴原点或上限位就绪 [-] / Z axis home or upper limit ready
    fPickZ        : LREAL := 0.0;      // 取料位下降目标 [毫米] / Pick position Z target
    fPlaceZ       : LREAL := 0.0;      // 放料位下降目标 [毫米] / Place position Z target
    fSafeZ        : LREAL := 50.0;     // 安全抬升位，用于抬升与中止 [毫米] / Safe lift height used for lifting and aborting
    fTravelX      : LREAL := 100.0;    // 取到放的横向行程 [毫米] / Horizontal travel from pick to place
    fSpeed        : LREAL := 200.0;    // 运动速度，域不小于 1 [毫米每秒] / Motion speed, not less than 1
    fAccel        : LREAL := 1000.0;   // 加减速度，域不小于 10 [毫米每二次方秒] / Acceleration and deceleration
    fPosTol       : LREAL := 0.5;      // 到位判定容差窗口 [毫米] / In-position tolerance window
    tGripTime     : TIME := T#200MS;   // 吸盘吸附建立时间 [毫秒] / Suction build-up time
    tBlowTime     : TIME := T#150MS;   // 破真空吹气时间 [毫秒] / Blow-off time
    tStepTimeout  : TIME := T#5S;      // 单步超时 [毫秒] / Per-step timeout
    tCycleTimeout : TIME := T#30S;     // 整循环超时，同时用作节拍秒表 [毫秒] / Whole-cycle timeout, also the cycle stopwatch
END_VAR
VAR_IN_OUT
    iAxisX        : I_DL_MotionAxis;      // X 轴接口引用，横向搬运 [-] / X axis interface reference
    iAxisY        : I_DL_MotionAxis;      // Y 轴接口引用，可选，未用时传同一实例 [-] / Y axis interface reference, optional
    iAxisZ        : I_DL_MotionAxis;      // Z 轴接口引用，升降 [-] / Z axis interface reference
    iVacuum       : I_DL_VacuumGenerator; // 真空发生器接口引用 [-] / Vacuum generator interface reference
END_VAR
VAR_OUTPUT
    eState        : E_DL_SpState;   // 工站状态，对外可观测 [-] / Station state, observable from outside
    nStepNo       : INT;            // 当前步号，1 到 9，0 为无常驻步 [步] / Current step number, 1 to 9, zero when idle
    bCycleDone    : BOOL;           // 单件循环完成，单拍脉冲 [-] / Cycle finished, single-cycle pulse
    bCycleOk      : BOOL;           // 本件合格，保持到下一件开始 [-] / Part accepted, held until the next cycle starts
    bPartLost     : BOOL;           // 搬运中真空丢失，保持 [-] / Part lost during transport, holding
    bError        : BOOL;           // 故障锁存 [-] / Fault latch
    uErrorId      : UDINT;          // 事件码，0 = 无事件 / Event code, 0 = no event
    tCycleTime    : TIME;           // 上一件节拍 [毫秒] / Cycle time of the last part
    tCycleTimeAvg : TIME;           // 节拍移动平均，八件窗 [毫秒] / Moving average over an eight-part window
    nOkCnt        : UDINT;          // 合格计数 [件] / Accepted part counter
    nNgCnt        : UDINT;          // 不合格计数 [件] / Rejected part counter
    bCallAndon    : BOOL;           // 需人工介入，供安灯系统消费 [-] / Manual intervention request for the andon system
END_VAR
VAR
    fbTrigStart   : R_TRIG;         // 启动沿检测，CASE 之外无条件刷新 [-] / Rising edge detector for the start input
    fbTrigReset   : R_TRIG;         // 复位沿检测，CASE 之外无条件刷新 [-] / Rising edge detector for the reset input
    fbStepTmo     : TON;            // 单步超时，CASE 之外无条件刷新 [-] / Per-step timeout timer
    fbCycleTmo    : TON;            // 整循环超时兼节拍秒表，CASE 之外无条件刷新 [-] / Cycle timeout and stopwatch timer
    fbGrip        : TON;            // 吸附建立计时 [-] / Suction build-up timer
    fbBlow        : TON;            // 破真空计时 [-] / Blow-off timer
    bInit         : BOOL := FALSE;  // 首扫标志，初值 FALSE，判据 NOT bInit（R19 范式）[-] / First-scan flag
    _eState       : E_DL_SpState := E_DL_SpState.eIdle;  // 内部状态机 [-] / Internal state machine
    nStep         : INT := 0;       // 内部步号，0 表示无常驻步 [步] / Internal step number
    nAbortStep    : INT := 0;       // 中止收尾子步，1 抬 Z，2 破真空，3 收口 [步] / Abort sub-step
    bStepActive   : BOOL;           // 本步已下发动作，防重复下发 [-] / TRUE once the current step has issued its action
    anCycleHistMs : ARRAY[0..7] OF DINT;  // 节拍历史窗，八件毫秒整数 [毫秒] / Cycle history window in milliseconds
    nHistIdx      : INT := 0;       // 历史窗写指针 [索引] / History write index
    nHistCnt      : INT := 0;       // 历史窗有效个数 [件] / Valid entries in the history window
    bStepTmoIn    : BOOL;           // 单步超时输入条件，先算后调 [-] / Step timer input condition
    bCycleTmoIn   : BOOL;           // 整循环超时输入条件，先算后调 [-] / Cycle timer input condition
    bGripIn       : BOOL;           // 吸附计时输入条件，先算后调 [-] / Grip timer input condition
    bBlowIn       : BOOL;           // 吹气计时输入条件，先算后调 [-] / Blow timer input condition
    tStepTmoUse   : TIME := T#5S;   // 生效单步超时（已钳位）[毫秒] / Effective step timeout
    tCycleTmoUse  : TIME := T#30S;  // 生效整循环超时（已钳位）[毫秒] / Effective cycle timeout
    tGripUse      : TIME := T#200MS; // 生效吸附时间（已钳位）[毫秒] / Effective grip time
    tBlowUse      : TIME := T#150MS; // 生效吹气时间（已钳位）[毫秒] / Effective blow time
    bAxisValid    : BOOL;           // 四个接口引用全部有效 [-] / TRUE when every injected interface is valid
    bFaultStopDone: BOOL;           // 进故障时轴停止指令已发过，防每拍重发 [-] / TRUE once the axes have been stopped on fault entry
    diCycleMs     : DINT;           // 本件节拍毫秒整数 [毫秒] / Cycle time in milliseconds
    diSumMs       : DINT;           // 窗口求和中间量 [毫秒] / Window sum
    i             : INT;            // 历史窗求和循环索引 [索引] / Summation index
    fSpeedUse     : REAL;           // 生效速度（已转为接口类型）[毫米每秒] / Effective speed converted for the interface
    fAccelUse     : REAL;           // 生效加速度（已转为接口类型）[毫米每二次方秒] / Effective acceleration converted for the interface
END_VAR
VAR CONSTANT
    DL_STEP_NUM    : INT   := 9;           // 总步数 [步] / Total step count
    DL_HIST_LEN    : INT   := 8;           // 节拍历史窗长度 [件] / Cycle history window length
    DL_SPEED_MIN   : LREAL := 1.0;         // 速度下限 [毫米每秒] / Speed lower bound
    DL_ACCEL_MIN   : LREAL := 10.0;        // 加速度下限 [毫米每二次方秒] / Acceleration lower bound
    DL_TMO_MAX     : TIME  := T#60S;       // 超时上限 [毫秒] / Timeout upper bound
    DL_GRIP_MAX    : TIME  := T#10S;       // 吸附与吹气时间上限 [毫秒] / Grip and blow time upper bound
    DL_POS_DEFAULT : LREAL := 50.0;        // 安全位兜底高度 [毫米] / Safe height fallback
    DL_AXIS_TOL_MIN: LREAL := 0.01;        // 到位容差下限 [毫米] / Minimum in-position tolerance
END_VAR

(*------------------------------------------------------------------------------
 * 段 1｜单拍输出预清零（R25 律①）
 *      Single-cycle output pre-clear
 *-----------------------------------------------------------------------------*)
bCycleDone := FALSE;

(*------------------------------------------------------------------------------
 * 段 2｜超时参数钳位（先钳位再调用，杜绝分支内调用实例）
 *      Timeout parameters clamped before the unconditional timer calls
 *-----------------------------------------------------------------------------*)
tStepTmoUse := tStepTimeout;
IF tStepTmoUse > DL_TMO_MAX THEN
    tStepTmoUse := DL_TMO_MAX;
ELSIF tStepTmoUse < T#10MS THEN
    tStepTmoUse := T#10MS;
END_IF

tCycleTmoUse := tCycleTimeout;
IF tCycleTmoUse > DL_TMO_MAX THEN
    tCycleTmoUse := DL_TMO_MAX;
ELSIF tCycleTmoUse < T#10MS THEN
    tCycleTmoUse := T#10MS;
END_IF

tGripUse := tGripTime;
IF tGripUse > DL_GRIP_MAX THEN
    tGripUse := DL_GRIP_MAX;
ELSIF tGripUse < T#0S THEN
    tGripUse := T#0S;
END_IF

tBlowUse := tBlowTime;
IF tBlowUse > DL_GRIP_MAX THEN
    tBlowUse := DL_GRIP_MAX;
ELSIF tBlowUse < T#0S THEN
    tBlowUse := T#0S;
END_IF

(*------------------------------------------------------------------------------
 * 段 3｜沿与定时器无条件刷新（R7 红线）：六个实例全部在 CASE 之外
 *      All six instances refreshed outside the CASE, mandatory by the red line
 *-----------------------------------------------------------------------------*)
fbTrigStart(CLK := bStart);
fbTrigReset(CLK := bReset);

IF bStepActive AND (_eState = E_DL_SpState.eExecute) THEN
    bStepTmoIn := TRUE;
ELSE
    bStepTmoIn := FALSE;
END_IF
fbStepTmo(IN := bStepTmoIn, PT := tStepTmoUse);

IF _eState = E_DL_SpState.eExecute THEN
    bCycleTmoIn := TRUE;
ELSE
    bCycleTmoIn := FALSE;
END_IF
fbCycleTmo(IN := bCycleTmoIn, PT := tCycleTmoUse);

IF bStepActive AND (nStep = 4) THEN
    bGripIn := TRUE;
ELSE
    bGripIn := FALSE;
END_IF
fbGrip(IN := bGripIn, PT := tGripUse);

IF bStepActive AND (nStep = 8) THEN
    bBlowIn := TRUE;
ELSE
    bBlowIn := FALSE;
END_IF
fbBlow(IN := bBlowIn, PT := tBlowUse);

(*------------------------------------------------------------------------------
 * 段 4｜首扫初始化（R19 唯一合法范式）
 *      First-scan initialisation with the canonical R19 pattern
 *-----------------------------------------------------------------------------*)
IF NOT bInit THEN
    _eState        := E_DL_SpState.eIdle;
    nStep          := 0;
    nAbortStep     := 0;
    bStepActive    := FALSE;
    nOkCnt         := 0;
    nNgCnt         := 0;
    nHistIdx       := 0;
    nHistCnt       := 0;
    bCycleOk       := FALSE;
    bPartLost      := FALSE;
    bError         := FALSE;
    uErrorId       := 16#0000_0000;
    bCallAndon     := FALSE;
    tCycleTime     := T#0S;
    tCycleTimeAvg  := T#0S;
    bFaultStopDone := FALSE;
    FOR i := 0 TO (DL_HIST_LEN - 1) DO
        anCycleHistMs[i] := 0;
    END_FOR
    bInit := TRUE;                       // 首扫只做一次
END_IF

(*------------------------------------------------------------------------------
 * 段 5｜接口有效性与运动参数兜底（接口引用未注入时不得动作）
 *      Interface validity and motion parameter fallback
 *-----------------------------------------------------------------------------*)
IF (iAxisX = 0) OR (iAxisZ = 0) OR (iVacuum = 0) THEN
    bAxisValid := FALSE;
ELSE
    bAxisValid := TRUE;
END_IF

IF fSpeed < DL_SPEED_MIN THEN
    fSpeedUse := LREAL_TO_REAL(DL_SPEED_MIN);
ELSE
    fSpeedUse := LREAL_TO_REAL(fSpeed);
END_IF

IF fAccel < DL_ACCEL_MIN THEN
    fAccelUse := LREAL_TO_REAL(DL_ACCEL_MIN);
ELSE
    fAccelUse := LREAL_TO_REAL(fAccel);
END_IF

(*------------------------------------------------------------------------------
 * 段 6｜前置安全（每拍最先判）：中止优先，其次保持
 *      Pre-emptive safety evaluation: abort first, then hold
 *-----------------------------------------------------------------------------*)
IF bAbort THEN
    IF (_eState <> E_DL_SpState.eFault) AND (_eState <> E_DL_SpState.eAborting) THEN
        nAbortStep  := 1;
        bStepActive := FALSE;
        _eState     := E_DL_SpState.eAborting;
    END_IF
END_IF

IF bHold AND (_eState = E_DL_SpState.eExecute) AND (NOT bStepActive) THEN
    _eState := E_DL_SpState.eHolding;
END_IF

(*------------------------------------------------------------------------------
 * 段 7｜主状态机（ENUM 加 CASE，含 ELSE 兜底）
 *      Main state machine with an ELSE fallback branch
 *-----------------------------------------------------------------------------*)
CASE _eState OF
    E_DL_SpState.eIdle:
        IF fbTrigStart.Q AND bEnable AND bAxisValid THEN
            bCycleOk := FALSE;                 // 新件开始，清上一件结论
            _eState   := E_DL_SpState.eStarting;
        END_IF

    E_DL_SpState.eStarting:
        (* 自检：Z 原点就绪、放料位空闲、取料位有件；缺一即业务态退回 *)
        IF bZHomeOk AND bPlaceClear AND bPartPresent THEN
            nStep       := 1;
            bStepActive := FALSE;
            bCallAndon  := FALSE;
            uErrorId    := 16#0000_0000;
            _eState     := E_DL_SpState.eExecute;
        ELSE
            bCallAndon := TRUE;                // 缺料或放料位占用：叫料，不锁故障
            uErrorId   := 16#0005_01B2;
            _eState    := E_DL_SpState.eIdle;
        END_IF

    E_DL_SpState.eExecute:
        (* 执行态本体在段 8 至段 11 中处理（步超时、动作下发、完成推进、循环超时）
           本分支必须显式列出：CASE 缺该标签会让 eExecute 落入 ELSE 兜底而被判为
           非法状态并锁故障，工站将永远无法执行。禁止在此分支内写任何动作。 *)

    E_DL_SpState.eHolding:
        (* 单拍过渡态：目的只是把进入动作与停留态分开，便于 HMI 看到一次跃迁 *)
        _eState := E_DL_SpState.eHeld;

    E_DL_SpState.eHeld:
        (* 已保持：不发任何运动指令，真空状态保持；释放后从当前步继续 *)
        IF NOT bHold THEN
            _eState := E_DL_SpState.eExecute;
        END_IF

    E_DL_SpState.eAborting:
        (* 中止收尾：逐拍推进，一个扫描周期只发一条指令 *)
        IF nAbortStep = 1 THEN
            iAxisZ.MoveAbsolute(fPos := LREAL_TO_REAL(fSafeZ), fVel := fSpeedUse, fAcc := fAccelUse);
            nAbortStep := 2;
        ELSIF nAbortStep = 2 THEN
            iVacuum.CmdBlowOff();
            nAbortStep := 3;
        ELSE
            nAbortStep  := 0;
            nStep       := 0;
            bStepActive := FALSE;
            uErrorId    := 16#0005_01B3;       // 信息级：正常中止完成
            _eState     := E_DL_SpState.eIdle;
        END_IF

    E_DL_SpState.eFault:
        nStep       := 0;
        bStepActive := FALSE;
        IF fbTrigReset.Q THEN
            bError         := FALSE;
            bPartLost      := FALSE;
            bCallAndon     := FALSE;
            uErrorId       := 16#0000_0000;
            bFaultStopDone := FALSE;
            _eState        := E_DL_SpState.eIdle;
        END_IF

    ELSE
        (* 非法枚举值兜底 *)
        _eState     := E_DL_SpState.eFault;
        uErrorId    := 16#0005_02B7;
        bError      := TRUE;
        nStep       := 0;
        bStepActive := FALSE;
END_CASE

(*------------------------------------------------------------------------------
 * 段 8｜执行态步序：单步超时监视
 *      Execute state, per-step timeout supervision
 *-----------------------------------------------------------------------------*)
IF (_eState = E_DL_SpState.eExecute) AND fbStepTmo.Q THEN
    IF nStep = 1 THEN
        uErrorId    := 16#0005_01B0;        // 原点未就绪：信息级，重试本步
        bStepActive := FALSE;
    ELSE
        CASE nStep OF
            2: uErrorId := 16#0005_02B0;
            3: uErrorId := 16#0005_02B1;
            5: uErrorId := 16#0005_02B2;
            6: uErrorId := 16#0005_02B3;
            7: uErrorId := 16#0005_02B4;
            8: uErrorId := 16#0005_02B5;
            9: uErrorId := 16#0005_02B6;
            ELSE
                uErrorId := 16#0005_02B7;
        END_CASE
        bError      := TRUE;
        bStepActive := FALSE;
        _eState     := E_DL_SpState.eFault;
    END_IF
END_IF

(*------------------------------------------------------------------------------
 * 段 9｜执行态步序：动作下发（每步只发一次）
 *      Execute state, action dispatch once per step
 *-----------------------------------------------------------------------------*)
IF (_eState = E_DL_SpState.eExecute) AND (NOT bStepActive) THEN
    CASE nStep OF
        1:
            (* 步 1：只确认原点，无下发动作；残留信息码已在 eStarting 自检通过时
               清零（段 7），此处绝不可再写 uErrorId := 0，否则本步超时码 01B0
               会被同拍覆盖，现场看不到「原点未就绪」的直接提示 *)
        2:
            iAxisX.MoveAbsolute(fPos := 0.0, fVel := fSpeedUse, fAcc := fAccelUse);
        3:
            iAxisZ.MoveAbsolute(fPos := LREAL_TO_REAL(fPickZ), fVel := fSpeedUse, fAcc := fAccelUse);
        4:
            iVacuum.CmdEvacuate();           // 开始抽真空
        5:
            iAxisZ.MoveAbsolute(fPos := LREAL_TO_REAL(fSafeZ), fVel := fSpeedUse, fAcc := fAccelUse);
        6:
            iAxisX.MoveAbsolute(fPos := LREAL_TO_REAL(fTravelX), fVel := fSpeedUse, fAcc := fAccelUse);
        7:
            iAxisZ.MoveAbsolute(fPos := LREAL_TO_REAL(fPlaceZ), fVel := fSpeedUse, fAcc := fAccelUse);
        8:
            iVacuum.CmdBlowOff();            // 破真空
        9:
            iAxisZ.MoveAbsolute(fPos := LREAL_TO_REAL(fSafeZ), fVel := fSpeedUse, fAcc := fAccelUse);
            iAxisX.MoveAbsolute(fPos := 0.0, fVel := fSpeedUse, fAcc := fAccelUse);
        ELSE
            bError   := TRUE;
            uErrorId := 16#0005_02B7;
            _eState  := E_DL_SpState.eFault;
    END_CASE
    bStepActive := TRUE;
END_IF

(*------------------------------------------------------------------------------
 * 段 10｜执行态步序：完成条件判定与推进
 *      Execute state, completion predicates and step advance
 *-----------------------------------------------------------------------------*)
IF (_eState = E_DL_SpState.eExecute) AND bStepActive THEN
    CASE nStep OF
        1:
            IF bZHomeOk THEN
                nStep       := 2;
                bStepActive := FALSE;
            END_IF
        2:
            IF (iAxisX.eState = E_DL_AxisState.eStandstill) AND
               (ABS(REAL_TO_LREAL(iAxisX.fPosition)) <= MAX(fPosTol, DL_AXIS_TOL_MIN)) THEN
                nStep       := 3;
                bStepActive := FALSE;
            END_IF
        3:
            IF (iAxisZ.eState = E_DL_AxisState.eStandstill) AND
               (ABS(REAL_TO_LREAL(iAxisZ.fPosition) - fPickZ) <= MAX(fPosTol, DL_AXIS_TOL_MIN)) THEN
                nStep       := 4;
                bStepActive := FALSE;
            END_IF
        4:
            IF fbGrip.Q THEN
                IF bVacuumOk THEN
                    nStep       := 5;                  // 吸附建立成功
                    bStepActive := FALSE;
                ELSE
                    (* 真空未建立：本件判 NG，叫料，回步 1，不锁故障 *)
                    nNgCnt     := nNgCnt + 1;
                    bCallAndon := TRUE;
                    uErrorId   := 16#0005_01B1;
                    iVacuum.CmdStop();
                    nStep       := 1;
                    bStepActive := FALSE;
                END_IF
            END_IF
        5:
            IF (iAxisZ.eState = E_DL_AxisState.eStandstill) AND
               (ABS(REAL_TO_LREAL(iAxisZ.fPosition) - fSafeZ) <= MAX(fPosTol, DL_AXIS_TOL_MIN)) THEN
                nStep       := 6;
                bStepActive := FALSE;
            END_IF
        6:
            IF (iAxisX.eState = E_DL_AxisState.eStandstill) AND
               (ABS(REAL_TO_LREAL(iAxisX.fPosition) - fTravelX) <= MAX(fPosTol, DL_AXIS_TOL_MIN)) THEN
                nStep       := 7;
                bStepActive := FALSE;
            END_IF
        7:
            IF NOT bVacuumOk THEN
                (* 搬运中掉件：故障级，转中止收尾，避免二次撞机 *)
                bPartLost := TRUE;
                uErrorId  := 16#0005_02B4;
                bError    := TRUE;
                nAbortStep  := 1;
                bStepActive := FALSE;
                _eState     := E_DL_SpState.eAborting;
            ELSIF (iAxisZ.eState = E_DL_AxisState.eStandstill) AND
                  (ABS(REAL_TO_LREAL(iAxisZ.fPosition) - fPlaceZ) <= MAX(fPosTol, DL_AXIS_TOL_MIN)) THEN
                nStep       := 8;
                bStepActive := FALSE;
            END_IF
        8:
            IF fbBlow.Q THEN
                nStep       := 9;
                bStepActive := FALSE;
            END_IF
        9:
            IF (iAxisX.eState = E_DL_AxisState.eStandstill) AND
               (ABS(REAL_TO_LREAL(iAxisX.fPosition)) <= MAX(fPosTol, DL_AXIS_TOL_MIN)) AND
               (iAxisZ.eState = E_DL_AxisState.eStandstill) AND
               (ABS(REAL_TO_LREAL(iAxisZ.fPosition) - fSafeZ) <= MAX(fPosTol, DL_AXIS_TOL_MIN)) THEN
                (* 单件结算：完成脉冲单拍，节拍入窗并重算平均 *)
                bCycleDone := TRUE;
                nOkCnt     := nOkCnt + 1;
                bCycleOk   := TRUE;
                tCycleTime := fbCycleTmo.ET;
                diCycleMs  := TIME_TO_DINT(tCycleTime);
                anCycleHistMs[nHistIdx] := diCycleMs;
                nHistIdx   := (nHistIdx + 1) MOD DL_HIST_LEN;
                IF nHistCnt < DL_HIST_LEN THEN
                    nHistCnt := nHistCnt + 1;
                END_IF
                diSumMs := 0;
                FOR i := 0 TO (nHistCnt - 1) DO
                    diSumMs := diSumMs + anCycleHistMs[i];
                END_FOR
                IF nHistCnt > 0 THEN
                    tCycleTimeAvg := DINT_TO_TIME(diSumMs / nHistCnt);
                END_IF
                nStep       := 0;
                bStepActive := FALSE;
                _eState     := E_DL_SpState.eIdle;
            END_IF
        ELSE
            bError   := TRUE;
            uErrorId := 16#0005_02B7;
            _eState  := E_DL_SpState.eFault;
    END_CASE
END_IF

(*------------------------------------------------------------------------------
 * 段 11｜整循环超时（业务保护）：执行态超时即转中止收尾，不直接锁故障
 *      Cycle timeout protection, aborts instead of latching a fault
 *-----------------------------------------------------------------------------*)
IF (_eState = E_DL_SpState.eExecute) AND fbCycleTmo.Q THEN
    uErrorId    := 16#0005_02B7;   // 循环超时复用兜底码，理由见头注释偏离登记 D3
    nAbortStep  := 1;
    bStepActive := FALSE;
    _eState     := E_DL_SpState.eAborting;
END_IF

(*------------------------------------------------------------------------------
 * 段 12｜进故障时的轴停止（只发一次，禁止每拍重发）
 *      Stop the axes once on fault entry, never re-issued every cycle
 *-----------------------------------------------------------------------------*)
IF (_eState = E_DL_SpState.eFault) AND (NOT bFaultStopDone) THEN
    (* 逐个判空再调用：Y 轴为可选注入，未注入时接口引用为 0，直接调用会落到
       空引用上产生未定义行为。bAxisValid 只覆盖 X / Z / 真空三路，不足以
       保护 Y 轴，故此处对四路一律显式判空，绝不依赖组态纪律。 *)
    IF iAxisX <> 0 THEN
        iAxisX.Stop();
    END_IF
    IF iAxisY <> 0 THEN
        iAxisY.Stop();
    END_IF
    IF iAxisZ <> 0 THEN
        iAxisZ.Stop();
    END_IF
    IF iVacuum <> 0 THEN
        iVacuum.CmdStop();
    END_IF
    bFaultStopDone := TRUE;
END_IF

(*------------------------------------------------------------------------------
 * 段 13｜输出每拍重写（R27）
 *      Outputs rewritten every cycle
 *-----------------------------------------------------------------------------*)
eState  := _eState;
nStepNo := nStep;

IF _eState = E_DL_SpState.eFault THEN
    bError := TRUE;
END_IF

(*------------------------------------------------------------------------------
 * 现场提示：
 *   1 步 1 走的是「确认原点就绪」而不是「回原点」：回原序列由
 *     FB_DL_AxisHomingSeq 承担，工站不做回原，避免两处在同一轴上写指令；
 *   2 保持态释放后从当前步继续，若保持发生在步 3 的下降途中，释放后不会
 *     重发下降指令，轴会继续走完原指令，这是刻意的（重发会造成指令覆盖）；
 *   3 节拍秒表用整循环超时定时器的已历时值，该定时器进执行态开始计时、
 *     离开执行态清零，故单件节拍不含待机等待时间。
 *-----------------------------------------------------------------------------*)
END_FUNCTION_BLOCK
